(* IEC 61131-3 sources: PortalRobot/Portal_robot/Device/application (part 2) *)

(* ---- PLC_PRG.ReadIoOverrides.st ---- *)
METHOD PRIVATE ReadIoOverrides

// --- BEGIN IMPLEMENTATION ---

udiIoNowMs := TIME_TO_UDINT(TIME());
IF NOT xIoInitialized THEN
    GVL_HMI.udiIoBootCounter := GVL_HMI.udiIoBootCounter + UDINT#1;
    IF GVL_HMI.udiIoBootCounter = UDINT#0 THEN GVL_HMI.udiIoBootCounter := UDINT#1; END_IF;
    udiIoLastTickMs := udiIoNowMs;
    // Старый запрос после перезапуска не должен исполняться сам собой.
    GVL_HMI.udiIoOverrideAckSeq := GVL_HMI.udiIoOverrideCommandSeq;
    GVL_HMI.udiIoEmergencyAckSeq := GVL_HMI.udiIoEmergencyCommandSeq;
END_IF;
IF udiIoNowMs >= udiIoLastTickMs THEN
    uliIoClockMs := uliIoClockMs + UDINT_TO_ULINT(udiIoNowMs - udiIoLastTickMs);
ELSE
    uliIoClockMs := uliIoClockMs + ULINT#4294967296 - UDINT_TO_ULINT(udiIoLastTickMs) + UDINT_TO_ULINT(udiIoNowMs);
END_IF;
udiIoLastTickMs := udiIoNowMs;
GVL_HMI.sIoClockMs := ULINT_TO_STRING(uliIoClockMs);

tonIoOverrideWatchdog(IN := GVL_HMI.udiIoOverrideHeartbeat = udiIoHeartbeatSeen, PT := T#3S);
IF GVL_HMI.udiIoOverrideHeartbeat <> udiIoHeartbeatSeen THEN
    udiIoHeartbeatSeen := GVL_HMI.udiIoOverrideHeartbeat;
END_IF;
IF udiIoNowMs >= GVL_HMI.udiIoOverrideHeartbeatAtMs THEN
    uliIoLeaseAgeMs := UDINT_TO_ULINT(udiIoNowMs) - UDINT_TO_ULINT(GVL_HMI.udiIoOverrideHeartbeatAtMs);
ELSE
    uliIoLeaseAgeMs := ULINT#4294967296 + UDINT_TO_ULINT(udiIoNowMs) - UDINT_TO_ULINT(GVL_HMI.udiIoOverrideHeartbeatAtMs);
END_IF;

xIoBusy := GVL_CELL_MANAGER.Status.xRunning OR GVL_CELL_MANAGER.Status.xBusy
    OR GVL_CELL_MANAGER.Status.xStopPending OR GVL_ROBOT.Status.xBusy
    OR xMotionBusy OR xGroupMotionBusy OR xPointCheckActive OR xPointCheckRequest
    OR xPowerTransitionActive OR SIMULATION_DYNAMICS.xBusy
    OR GVL_HMI.xRobotManualExecute OR GVL_HMI.stRobotCommand.xExecute
    OR GVL_CELL_CONTROL.xStart
    OR (GVL_HMI.udiTwinCommandSeq <> GVL_HMI.udiTwinAckSeq);
// Реальный цикл станка нельзя скрыть подменой его DI.
IF xPhysicalNormal AND GVL_PHYSICAL_IO.xMappingVerified THEN
    xIoBusy := xIoBusy OR GVL_PHYSICAL_IO.xDiMachine1CycleActive
        OR GVL_PHYSICAL_IO.xDiMachine2CycleActive OR GVL_PHYSICAL_IO.xDiMachine3CycleActive;
END_IF;
FOR uiIoIndex := UINT#1 TO UINT#3 DO
    xIoBusy := xIoBusy OR GVL_MACHINE.Status[uiIoIndex].xBusy OR GVL_MACHINE.Status[uiIoIndex].xProcessing
        OR GVL_HMI.axMachineManualHatchOpen[uiIoIndex] OR GVL_HMI.axMachineManualHatchClose[uiIoIndex]
        OR GVL_HMI.axMachineManualHatchUnlock[uiIoIndex] OR GVL_HMI.axMachineManualHatchLock[uiIoIndex]
        OR GVL_HMI.axMachineManualChuckOpen[uiIoIndex] OR GVL_HMI.axMachineManualChuckClose[uiIoIndex]
        OR GVL_HMI.astAxisHmiCommand[uiIoIndex].xJogPositive
        OR GVL_HMI.astAxisHmiCommand[uiIoIndex].xJogNegative
        OR GVL_HMI.astAxisHmiCommand[uiIoIndex].xHome
        OR GVL_HMI.astAxisHmiCommand[uiIoIndex].xMoveAbsolute
        OR GVL_HMI.astAxisHmiCommand[uiIoIndex].xMoveRelative;
END_FOR;
FOR uiIoIndex := UINT#1 TO UINT#2 DO
    xIoBusy := xIoBusy OR GVL_MAGAZINE.astStatus[uiIoIndex].xBusy
        OR GVL_TWO_PALLET.astStatus[uiIoIndex].xBusy;
END_FOR;
// Ручной режим сигналов включается одним запросом. Технологических допусков здесь нет.
xIoManualEndedByOperator := FALSE;
IF xIoManualActive AND (NOT GVL_CELL_CONTROL.xManual OR NOT xHmiConnectionAlive
    OR CONTROLLER_DIAGNOSTICS.Status.xAlarmActive
    OR tonIoOverrideWatchdog.Q OR (uliIoLeaseAgeMs > ULINT#3000)
    OR ((GVL_HMI.udiCellModeCommandSeq <> GVL_HMI.udiCellModeAckSeq) AND NOT GVL_HMI.xCellManualRequest)) THEN
    xIoManualActive := FALSE;
END_IF;
// Прямой ручной слой доступен и при зависших Busy/Processing владельцев.
// Их задания отменяются при передаче управления; xIoBusy остаётся диагностикой
// и условием снятия отдельного программного аварийного останова.
GVL_HMI.xIoManualStartAllowed := GVL_CELL_CONTROL.xManual AND NOT xIoManualActive
    AND NOT CONTROLLER_DIAGNOSTICS.Status.xAlarmActive
    AND NOT ((GVL_HMI.udiCellModeCommandSeq <> GVL_HMI.udiCellModeAckSeq) AND NOT GVL_HMI.xCellManualRequest);
xIoOverrideRejected := FALSE;
udiIoRequestSeq := GVL_HMI.udiIoOverrideCommandSeq;
uiIoRequestAction := GVL_HMI.uiIoOverrideAction;
uiIoRequestIndex := GVL_HMI.uiIoOverrideIndex;
xIoRequestValue := GVL_HMI.xIoOverrideValue;
IF udiIoRequestSeq <> GVL_HMI.udiIoOverrideAckSeq THEN
    IF (uiIoRequestAction = UINT#8) OR (uiIoRequestAction = UINT#9) OR (uiIoRequestAction = UINT#7) THEN
        GVL_HMI.uiIoOverrideResult := UINT#4;
        IF IsHmiCommandFresh(udiIssuedAtMs := GVL_HMI.udiIoOverrideIssuedAtMs) THEN
            GVL_HMI.uiIoOverrideResult := UINT#1;
            IF uiIoRequestAction = UINT#8 THEN
                IF NOT xHmiConnectionAlive OR tonIoOverrideWatchdog.Q OR (uliIoLeaseAgeMs > ULINT#3000) THEN
                    GVL_HMI.uiIoOverrideResult := UINT#4;
                ELSIF xIoManualActive THEN
                    // Повтор входа не перезаписывает уже выбранные ручные уровни.
                    GVL_HMI.uiIoOverrideResult := UINT#1;
                ELSIF GVL_HMI.xIoManualStartAllowed THEN
                    FOR uiIoIndex := UINT#1 TO UINT#50 DO
                        axIoDoForceValue[uiIoIndex] := axIoOutput[uiIoIndex];
                        axIoDoForced[uiIoIndex] := FALSE;
                    END_FOR;
                    xIoManualActive := TRUE;
                ELSE
                    GVL_HMI.uiIoOverrideResult := UINT#2;
                END_IF;
            ELSE
                xIoManualActive := FALSE;
                xIoManualEndedByOperator := TRUE;
            END_IF;
        END_IF;
        // Для входа/выхода из режима Ack выдаёт ApplyIoOutputOverrides после назначения DO.
    END_IF;
END_IF;

GVL_HMI.xIoManualControlActive := xIoManualActive;
GVL_HMI.xIoManualStartAllowed := GVL_HMI.xIoManualStartAllowed AND NOT xIoManualActive;
GVL_HMI.xIoOverrideAllowed := xIoManualActive AND GVL_CELL_CONTROL.xManual;
IF GVL_HMI.xIoOverrideAllowed THEN GVL_HMI.uiIoOverrideBlockReason := UINT#0;
ELSIF NOT GVL_CELL_CONTROL.xManual THEN GVL_HMI.uiIoOverrideBlockReason := UINT#2;
ELSE GVL_HMI.uiIoOverrideBlockReason := UINT#7;
END_IF;

IF NOT GVL_HMI.xIoOverrideAllowed THEN
    FOR uiIoIndex := UINT#1 TO UINT#84 DO
        IF axIoForced[uiIoIndex] THEN
            IF xIoManualEndedByOperator THEN
                AppendIoEvent(usiDirection := USINT#1, uiIndex := uiIoIndex, usiKind := USINT#5,
                    xOld := axIoForceValue[uiIoIndex], xNew := axIoRawDi[uiIoIndex]);
            ELSE
                AppendIoEvent(usiDirection := USINT#1, uiIndex := uiIoIndex, usiKind := USINT#6,
                    xOld := axIoForceValue[uiIoIndex], xNew := axIoRawDi[uiIoIndex]);
            END_IF;
            axIoForced[uiIoIndex] := FALSE;
        END_IF;
    END_FOR;
END_IF;

IF (udiIoRequestSeq <> GVL_HMI.udiIoOverrideAckSeq)
AND NOT ((uiIoRequestAction >= UINT#4) AND (uiIoRequestAction <= UINT#9)) THEN
    GVL_HMI.uiIoOverrideResult := UINT#3;
    IF NOT IsHmiCommandFresh(udiIssuedAtMs := GVL_HMI.udiIoOverrideIssuedAtMs) THEN
        GVL_HMI.uiIoOverrideResult := UINT#4;
    ELSIF uiIoRequestAction = UINT#3 THEN
        FOR uiIoIndex := UINT#1 TO UINT#84 DO
            IF axIoForced[uiIoIndex] THEN
                AppendIoEvent(usiDirection := USINT#1, uiIndex := uiIoIndex, usiKind := USINT#5,
                    xOld := axIoForceValue[uiIoIndex], xNew := axIoRawDi[uiIoIndex]);
                axIoForced[uiIoIndex] := FALSE;
            END_IF;
        END_FOR;
        GVL_HMI.uiIoOverrideResult := UINT#1;
    ELSIF (uiIoRequestIndex >= UINT#1) AND (uiIoRequestIndex <= UINT#84) THEN
        IF uiIoRequestAction = UINT#2 THEN
            IF axIoForced[uiIoRequestIndex] THEN
                AppendIoEvent(usiDirection := USINT#1, uiIndex := uiIoRequestIndex, usiKind := USINT#5,
                    xOld := axIoForceValue[uiIoRequestIndex], xNew := axIoRawDi[uiIoRequestIndex]);
                axIoForced[uiIoRequestIndex] := FALSE;
            END_IF;
            GVL_HMI.uiIoOverrideResult := UINT#1;
        ELSIF uiIoRequestAction = UINT#1 THEN
            IF GVL_HMI.xIoOverrideAllowed THEN
                IF NOT axIoForced[uiIoRequestIndex] OR (axIoForceValue[uiIoRequestIndex] <> xIoRequestValue) THEN
                    AppendIoEvent(usiDirection := USINT#1, uiIndex := uiIoRequestIndex, usiKind := USINT#4,
                        xOld := axPhysicalRaw[uiIoRequestIndex], xNew := xIoRequestValue);
                END_IF;
                axIoForced[uiIoRequestIndex] := TRUE;
                axIoForceValue[uiIoRequestIndex] := xIoRequestValue;
                GVL_HMI.uiIoOverrideResult := UINT#1;
            ELSE
                GVL_HMI.uiIoOverrideResult := UINT#2;
            END_IF;
        END_IF;
    END_IF;
    xIoOverrideRejected := GVL_HMI.uiIoOverrideResult <> UINT#1;
    GVL_HMI.udiIoOverrideAckSeq := udiIoRequestSeq;
END_IF;
FOR uiIoIndex := UINT#1 TO UINT#84 DO
    IF axIoForced[uiIoIndex] THEN axPhysicalRaw[uiIoIndex] := axIoForceValue[uiIoIndex]; END_IF;
END_FOR;

(* ---- PLC_PRG.ReadPhysicalInputs.st ---- *)
METHOD PRIVATE ReadPhysicalInputs

// --- BEGIN IMPLEMENTATION ---

// Единственная страница назначения входов. Сначала фильтры, затем технологические FB.
// Тестовые среды используют модели; сырые входы приводов ГК читает RunGeometryControl.
xPhysicalNormal := GVL_CELL_SETTINGS.eTestEnvironment = E_CELL_TEST_ENVIRONMENT.NORMAL;
GVL_PHYSICAL_IO.xNormalActive := xPhysicalNormal AND GVL_PHYSICAL_IO.xMappingVerified;
xPhysicalInputEnable := GVL_PHYSICAL_IO.xNormalActive;

axPhysicalRaw[1] := GVL_PHYSICAL_IO.xDiMachine1Ready;
axPhysicalRaw[2] := GVL_PHYSICAL_IO.xDiMachine1Alarm;
axPhysicalRaw[3] := GVL_PHYSICAL_IO.xDiMachine1DoorOpen;
axPhysicalRaw[4] := GVL_PHYSICAL_IO.xDiMachine1DoorClosed;
axPhysicalRaw[5] := GVL_PHYSICAL_IO.xDiMachine1HatchLocked;
axPhysicalRaw[6] := GVL_PHYSICAL_IO.xDiMachine1SafetyDoorOpen;
axPhysicalRaw[7] := GVL_PHYSICAL_IO.xDiMachine1SafetyDoorClosed;
axPhysicalRaw[8] := GVL_PHYSICAL_IO.xDiMachine1ChuckClamped;
axPhysicalRaw[9] := GVL_PHYSICAL_IO.xDiMachine1ChuckUnclamped;
axPhysicalRaw[10] := GVL_PHYSICAL_IO.xDiMachine1CycleActive;
axPhysicalRaw[11] := GVL_PHYSICAL_IO.xDiMachine1CycleDone;
axPhysicalRaw[12] := GVL_PHYSICAL_IO.xDiMachine2Ready;
axPhysicalRaw[13] := GVL_PHYSICAL_IO.xDiMachine2Alarm;
axPhysicalRaw[14] := GVL_PHYSICAL_IO.xDiMachine2DoorOpen;
axPhysicalRaw[15] := GVL_PHYSICAL_IO.xDiMachine2DoorClosed;
axPhysicalRaw[16] := GVL_PHYSICAL_IO.xDiMachine2HatchLocked;
axPhysicalRaw[17] := GVL_PHYSICAL_IO.xDiMachine2SafetyDoorOpen;
axPhysicalRaw[18] := GVL_PHYSICAL_IO.xDiMachine2SafetyDoorClosed;
axPhysicalRaw[19] := GVL_PHYSICAL_IO.xDiMachine2ChuckClamped;
axPhysicalRaw[20] := GVL_PHYSICAL_IO.xDiMachine2ChuckUnclamped;
axPhysicalRaw[21] := GVL_PHYSICAL_IO.xDiMachine2CycleActive;
axPhysicalRaw[22] := GVL_PHYSICAL_IO.xDiMachine2CycleDone;
axPhysicalRaw[23] := GVL_PHYSICAL_IO.xDiMachine3Ready;
axPhysicalRaw[24] := GVL_PHYSICAL_IO.xDiMachine3Alarm;
axPhysicalRaw[25] := GVL_PHYSICAL_IO.xDiMachine3DoorOpen;
axPhysicalRaw[26] := GVL_PHYSICAL_IO.xDiMachine3DoorClosed;
axPhysicalRaw[27] := GVL_PHYSICAL_IO.xDiMachine3HatchLocked;
axPhysicalRaw[28] := GVL_PHYSICAL_IO.xDiMachine3SafetyDoorOpen;
axPhysicalRaw[29] := GVL_PHYSICAL_IO.xDiMachine3SafetyDoorClosed;
axPhysicalRaw[30] := GVL_PHYSICAL_IO.xDiMachine3ChuckClamped;
axPhysicalRaw[31] := GVL_PHYSICAL_IO.xDiMachine3ChuckUnclamped;
axPhysicalRaw[32] := GVL_PHYSICAL_IO.xDiMachine3CycleActive;
axPhysicalRaw[33] := GVL_PHYSICAL_IO.xDiMachine3CycleDone;
axPhysicalRaw[34] := GVL_PHYSICAL_IO.xDiGripper1Open;
axPhysicalRaw[35] := GVL_PHYSICAL_IO.xDiGripper1Closed;
axPhysicalRaw[36] := GVL_PHYSICAL_IO.xDiGripper2Open;
axPhysicalRaw[37] := GVL_PHYSICAL_IO.xDiGripper2Closed;
axPhysicalRaw[38] := GVL_PHYSICAL_IO.xDiRotatedToBlank;
axPhysicalRaw[39] := GVL_PHYSICAL_IO.xDiRotatedToDetail;
axPhysicalRaw[40] := GVL_PHYSICAL_IO.xDiCellStartButtonInput;
axPhysicalRaw[41] := GVL_PHYSICAL_IO.xDiCellStopButtonInput;
axPhysicalRaw[42] := GVL_PHYSICAL_IO.xDiCellResetButtonInput;
axPhysicalRaw[43] := GVL_PHYSICAL_IO.xDiEmergencyStopStation1Ok;
axPhysicalRaw[44] := GVL_PHYSICAL_IO.xDiEmergencyStopStation2Ok;
axPhysicalRaw[45] := GVL_PHYSICAL_IO.xDiEmergencyStopStation3Ok;
axPhysicalRaw[46] := GVL_PHYSICAL_IO.xDiEmergencyStopStation4Ok;
axPhysicalRaw[47] := GVL_PHYSICAL_IO.xDiEmergencyStopCabinet1Ok;
axPhysicalRaw[48] := GVL_PHYSICAL_IO.xDiEmergencyStopCabinet2Ok;
axPhysicalRaw[49] := GVL_PHYSICAL_IO.xDiEmergencyStopMpgOk;
axPhysicalRaw[50] := GVL_PHYSICAL_IO.xDiDoor1LockClosed;
axPhysicalRaw[51] := GVL_PHYSICAL_IO.xDiDoor2LockClosed;
axPhysicalRaw[52] := GVL_PHYSICAL_IO.xDiDoor3LockClosed;
axPhysicalRaw[53] := GVL_PHYSICAL_IO.xDiDoor4LockClosed;
axPhysicalRaw[54] := GVL_PHYSICAL_IO.xDiSafetyRelayOkInput;
axPhysicalRaw[55] := GVL_PHYSICAL_IO.xDiPhaseRelayOkInput;
axPhysicalRaw[56] := GVL_PHYSICAL_IO.xDiPressureRelayOkInput;
axPhysicalRaw[57] := GVL_PHYSICAL_IO.xDiMpgAxisXInput;
axPhysicalRaw[58] := GVL_PHYSICAL_IO.xDiMpgAxisYInput;
axPhysicalRaw[59] := GVL_PHYSICAL_IO.xDiMpgAxisZInput;
axPhysicalRaw[60] := GVL_PHYSICAL_IO.xDiMpgMultiplier1Input;
axPhysicalRaw[61] := GVL_PHYSICAL_IO.xDiMpgMultiplier10Input;
axPhysicalRaw[62] := GVL_PHYSICAL_IO.xDiMpgMultiplier100Input;
axPhysicalRaw[63] := GVL_PHYSICAL_IO.xDiMagazine1LockIn;
axPhysicalRaw[64] := GVL_PHYSICAL_IO.xDiMagazine1LockOut;
axPhysicalRaw[65] := GVL_PHYSICAL_IO.xDiMagazine1StopIn;
axPhysicalRaw[66] := GVL_PHYSICAL_IO.xDiMagazine1StopOut;
axPhysicalRaw[67] := GVL_PHYSICAL_IO.xDiMagazine1LiftUp;
axPhysicalRaw[68] := GVL_PHYSICAL_IO.xDiMagazine1LiftDown;
axPhysicalRaw[69] := GVL_PHYSICAL_IO.xDiDoor1UnlockButton;
axPhysicalRaw[70] := GVL_PHYSICAL_IO.xDiDoor2UnlockButton;
axPhysicalRaw[71] := GVL_PHYSICAL_IO.xDiDoor3UnlockButton;
axPhysicalRaw[72] := GVL_PHYSICAL_IO.xDiDoor4UnlockButton;
axPhysicalRaw[73] := GVL_PHYSICAL_IO.xDiMagazine2LockIn;
axPhysicalRaw[74] := GVL_PHYSICAL_IO.xDiMagazine2LockOut;
axPhysicalRaw[75] := GVL_PHYSICAL_IO.xDiMagazine2StopIn;
axPhysicalRaw[76] := GVL_PHYSICAL_IO.xDiMagazine2StopOut;
axPhysicalRaw[77] := GVL_PHYSICAL_IO.xDiMagazine2LiftUp;
axPhysicalRaw[78] := GVL_PHYSICAL_IO.xDiMagazine2LiftDown;

axPhysicalRaw[79] := GVL_PHYSICAL_IO.xDiGk1PartAtEnd;
axPhysicalRaw[80] := GVL_PHYSICAL_IO.xDiGk2PartAtEnd;

axPhysicalRaw[81] := GVL_PHYSICAL_IO.xDiGk1DriveAlarm;
axPhysicalRaw[82] := GVL_PHYSICAL_IO.xDiGk1DriveRunning;
axPhysicalRaw[83] := GVL_PHYSICAL_IO.xDiGk2DriveAlarm;
axPhysicalRaw[84] := GVL_PHYSICAL_IO.xDiGk2DriveRunning;
// Клеммы сохраняются отдельно: ручная подмена не пишет в переменную I/O Mapping.
FOR uiIoIndex := UINT#1 TO UINT#84 DO
    axIoRawDi[uiIoIndex] := axPhysicalRaw[uiIoIndex];
END_FOR;
ReadIoOverrides();
FOR uiIoIndex := UINT#1 TO UINT#84 DO
    IF axIoForced[uiIoIndex] THEN
        axPhysicalRaw[uiIoIndex] := axIoForceValue[uiIoIndex];
    END_IF;
END_FOR;

FOR uiPhysicalInput := 1 TO 80 DO
	tPhysicalRise := GVL_CELL_SETTINGS.tInputFilterRise;
	tPhysicalFall := GVL_CELL_SETTINGS.tInputFilterFall;
	// Срабатывание опасного состояния не задерживается; восстановление фильтруется.
	CASE uiPhysicalInput OF
		2, 13, 24, 41:
			tPhysicalRise := T#0MS;
		1, 3, 4, 5, 6, 7, 8, 9, 12, 14, 15, 16, 17, 18, 19, 20, 23, 25, 26, 27, 28, 29, 30, 31, 34, 35, 36, 37, 38, 39, 43, 44, 45, 46, 47, 48, 49, 50, 51, 52, 53, 54, 55, 56, 63, 64, 65, 66, 67, 68, 73, 74, 75, 76, 77, 78, 79, 80:
			tPhysicalFall := T#0MS;
	END_CASE;
	xPhysicalInputEnable := xPhysicalNormal AND (GVL_PHYSICAL_IO.xMappingVerified OR axIoForced[uiPhysicalInput]);
	afbPhysicalInputFilter[uiPhysicalInput](
		xEnable := xPhysicalInputEnable, xInput := axPhysicalRaw[uiPhysicalInput],
		tRise := tPhysicalRise, tFall := tPhysicalFall);
	axPhysicalFiltered[uiPhysicalInput] := afbPhysicalInputFilter[uiPhysicalInput].xFiltered;
	IF NOT xPhysicalInputEnable THEN
		axPhysicalButtonArmed[uiPhysicalInput] := FALSE;
	ELSIF NOT axPhysicalRaw[uiPhysicalInput] THEN
		axPhysicalButtonArmed[uiPhysicalInput] := TRUE;
	END_IF;
END_FOR;

// Датчики используются FB_GEOMETRY_CONTROL; в NORMAL доступна диагностическая подмена до подтверждения карты.
GVL_PHYSICAL_IO.axGkPartAtEnd[1] := axPhysicalFiltered[79];
GVL_PHYSICAL_IO.axGkPartAtEnd[2] := axPhysicalFiltered[80];

IF xPhysicalNormal THEN
	GVL_MACHINE.astPhysicalInput[1].xReady := axPhysicalFiltered[1];
	GVL_MACHINE.astPhysicalInput[1].xAlarm := axPhysicalFiltered[2];
	GVL_MACHINE.astPhysicalInput[1].xDoorOpen := axPhysicalFiltered[3];
	GVL_MACHINE.astPhysicalInput[1].xDoorClosed := axPhysicalFiltered[4];
	GVL_MACHINE.astPhysicalInput[1].xHatchLocked := axPhysicalFiltered[5];
	GVL_MACHINE.astPhysicalInput[1].xSafetyDoorOpen := axPhysicalFiltered[6];
	GVL_MACHINE.astPhysicalInput[1].xSafetyDoorClosed := axPhysicalFiltered[7];
	GVL_MACHINE.astPhysicalInput[1].xChuckClamped := axPhysicalFiltered[8];
	GVL_MACHINE.astPhysicalInput[1].xChuckUnclamped := axPhysicalFiltered[9];
	GVL_MACHINE.astPhysicalInput[1].xCycleActive := axPhysicalFiltered[10];
	GVL_MACHINE.astPhysicalInput[1].xCycleDone := axPhysicalFiltered[11];
	GVL_MACHINE.astPhysicalInput[2].xReady := axPhysicalFiltered[12];
	GVL_MACHINE.astPhysicalInput[2].xAlarm := axPhysicalFiltered[13];
	GVL_MACHINE.astPhysicalInput[2].xDoorOpen := axPhysicalFiltered[14];
	GVL_MACHINE.astPhysicalInput[2].xDoorClosed := axPhysicalFiltered[15];
	GVL_MACHINE.astPhysicalInput[2].xHatchLocked := axPhysicalFiltered[16];
	GVL_MACHINE.astPhysicalInput[2].xSafetyDoorOpen := axPhysicalFiltered[17];
	GVL_MACHINE.astPhysicalInput[2].xSafetyDoorClosed := axPhysicalFiltered[18];
	GVL_MACHINE.astPhysicalInput[2].xChuckClamped := axPhysicalFiltered[19];
	GVL_MACHINE.astPhysicalInput[2].xChuckUnclamped := axPhysicalFiltered[20];
	GVL_MACHINE.astPhysicalInput[2].xCycleActive := axPhysicalFiltered[21];
	GVL_MACHINE.astPhysicalInput[2].xCycleDone := axPhysicalFiltered[22];
	GVL_MACHINE.astPhysicalInput[3].xReady := axPhysicalFiltered[23];
	GVL_MACHINE.astPhysicalInput[3].xAlarm := axPhysicalFiltered[24];
	GVL_MACHINE.astPhysicalInput[3].xDoorOpen := axPhysicalFiltered[25];
	GVL_MACHINE.astPhysicalInput[3].xDoorClosed := axPhysicalFiltered[26];
	GVL_MACHINE.astPhysicalInput[3].xHatchLocked := axPhysicalFiltered[27];
	GVL_MACHINE.astPhysicalInput[3].xSafetyDoorOpen := axPhysicalFiltered[28];
	GVL_MACHINE.astPhysicalInput[3].xSafetyDoorClosed := axPhysicalFiltered[29];
	GVL_MACHINE.astPhysicalInput[3].xChuckClamped := axPhysicalFiltered[30];
	GVL_MACHINE.astPhysicalInput[3].xChuckUnclamped := axPhysicalFiltered[31];
	GVL_MACHINE.astPhysicalInput[3].xCycleActive := axPhysicalFiltered[32];
	GVL_MACHINE.astPhysicalInput[3].xCycleDone := axPhysicalFiltered[33];
	GVL_PHYSICAL_IO.stGripperFeedback.xGripper1Open := axPhysicalFiltered[34];
	GVL_PHYSICAL_IO.stGripperFeedback.xGripper1Closed := axPhysicalFiltered[35];
	GVL_PHYSICAL_IO.stGripperFeedback.xGripper2Open := axPhysicalFiltered[36];
	GVL_PHYSICAL_IO.stGripperFeedback.xGripper2Closed := axPhysicalFiltered[37];
	GVL_PHYSICAL_IO.stGripperFeedback.xRotatedToBlank := axPhysicalFiltered[38];
	GVL_PHYSICAL_IO.stGripperFeedback.xRotatedToDetail := axPhysicalFiltered[39];
	GVL_CELL_SAFETY_IO.xCellStartButtonInput := axPhysicalFiltered[40] AND axPhysicalButtonArmed[40];
	GVL_CELL_SAFETY_IO.xCellStopButtonInput := axPhysicalFiltered[41];
	GVL_CELL_SAFETY_IO.xCellResetButtonInput := axPhysicalFiltered[42] AND axPhysicalButtonArmed[42];
	GVL_CELL_SAFETY_IO.axEmergencyStopButtonStationInput[1] := NOT axPhysicalFiltered[43];
	GVL_CELL_SAFETY_IO.axEmergencyStopButtonStationInput[2] := NOT axPhysicalFiltered[44];
	GVL_CELL_SAFETY_IO.axEmergencyStopButtonStationInput[3] := NOT axPhysicalFiltered[45];
	GVL_CELL_SAFETY_IO.axEmergencyStopButtonStationInput[4] := NOT axPhysicalFiltered[46];
	GVL_CELL_SAFETY_IO.axEmergencyStopCabinetInput[1] := NOT axPhysicalFiltered[47];
	GVL_CELL_SAFETY_IO.axEmergencyStopCabinetInput[2] := NOT axPhysicalFiltered[48];
	GVL_CELL_SAFETY_IO.xEmergencyStopMpgInput := NOT axPhysicalFiltered[49];
	GVL_CELL_SAFETY_IO.axDoorLockClosedInput[1] := axPhysicalFiltered[50];
	GVL_CELL_SAFETY_IO.axDoorLockClosedInput[2] := axPhysicalFiltered[51];
	GVL_CELL_SAFETY_IO.axDoorLockClosedInput[3] := axPhysicalFiltered[52];
	GVL_CELL_SAFETY_IO.axDoorLockClosedInput[4] := axPhysicalFiltered[53];
	GVL_CELL_SAFETY_IO.xSafetyRelayOkInput := axPhysicalFiltered[54];
	GVL_CELL_SAFETY_IO.xPhaseRelayOkInput := axPhysicalFiltered[55];
	GVL_CELL_SAFETY_IO.xPressureRelayOkInput := axPhysicalFiltered[56];
	GVL_CELL_SAFETY_IO.xMpgAxisXInput := axPhysicalFiltered[57];
	GVL_CELL_SAFETY_IO.xMpgAxisYInput := axPhysicalFiltered[58];
	GVL_CELL_SAFETY_IO.xMpgAxisZInput := axPhysicalFiltered[59];
	GVL_CELL_SAFETY_IO.xMpgMultiplier1Input := axPhysicalFiltered[60];
	GVL_CELL_SAFETY_IO.xMpgMultiplier10Input := axPhysicalFiltered[61];
	GVL_CELL_SAFETY_IO.xMpgMultiplier100Input := axPhysicalFiltered[62];
	GVL_TWO_PALLET.astInput[1].xLockIn := axPhysicalFiltered[63];
	GVL_TWO_PALLET.astInput[1].xLockOut := axPhysicalFiltered[64];
	GVL_TWO_PALLET.astInput[1].xStopIn := axPhysicalFiltered[65];
	GVL_TWO_PALLET.astInput[1].xStopOut := axPhysicalFiltered[66];
	GVL_TWO_PALLET.astInput[1].xLiftUp := axPhysicalFiltered[67];
	GVL_TWO_PALLET.astInput[1].xLiftDown := axPhysicalFiltered[68];
	GVL_CELL_SAFETY_IO.axDoorUnlockButtonInput[1] := axPhysicalFiltered[69] AND axPhysicalButtonArmed[69];
	GVL_CELL_SAFETY_IO.axDoorUnlockButtonInput[2] := axPhysicalFiltered[70] AND axPhysicalButtonArmed[70];
	GVL_CELL_SAFETY_IO.axDoorUnlockButtonInput[3] := axPhysicalFiltered[71] AND axPhysicalButtonArmed[71];
	GVL_CELL_SAFETY_IO.axDoorUnlockButtonInput[4] := axPhysicalFiltered[72] AND axPhysicalButtonArmed[72];
	GVL_TWO_PALLET.astInput[2].xLockIn := axPhysicalFiltered[73];
	GVL_TWO_PALLET.astInput[2].xLockOut := axPhysicalFiltered[74];
	GVL_TWO_PALLET.astInput[2].xStopIn := axPhysicalFiltered[75];
	GVL_TWO_PALLET.astInput[2].xStopOut := axPhysicalFiltered[76];
	GVL_TWO_PALLET.astInput[2].xLiftUp := axPhysicalFiltered[77];
	GVL_TWO_PALLET.astInput[2].xLiftDown := axPhysicalFiltered[78];
	GVL_TWO_PALLET.astInput[1].xIoMapped := GVL_PHYSICAL_IO.xNormalActive;
	GVL_TWO_PALLET.astInput[2].xIoMapped := GVL_PHYSICAL_IO.xNormalActive;
	GVL_MACHINE.astPhysicalInput[1].tRemaining := T#0MS;
	GVL_MACHINE.astPhysicalInput[2].tRemaining := T#0MS;
	GVL_MACHINE.astPhysicalInput[3].tRemaining := T#0MS;
ELSIF xPhysicalWasNormal THEN
	GVL_CELL_SAFETY_IO.xCellStartButtonInput := FALSE;
	GVL_CELL_SAFETY_IO.xCellStopButtonInput := FALSE;
	GVL_CELL_SAFETY_IO.xCellResetButtonInput := FALSE;
	GVL_CELL_SAFETY_IO.axEmergencyStopButtonStationInput[1] := FALSE;
	GVL_CELL_SAFETY_IO.axEmergencyStopButtonStationInput[2] := FALSE;
	GVL_CELL_SAFETY_IO.axEmergencyStopButtonStationInput[3] := FALSE;
	GVL_CELL_SAFETY_IO.axEmergencyStopButtonStationInput[4] := FALSE;
	GVL_CELL_SAFETY_IO.axEmergencyStopCabinetInput[1] := FALSE;
	GVL_CELL_SAFETY_IO.axEmergencyStopCabinetInput[2] := FALSE;
	GVL_CELL_SAFETY_IO.xEmergencyStopMpgInput := FALSE;
	GVL_CELL_SAFETY_IO.axDoorLockClosedInput[1] := TRUE;
	GVL_CELL_SAFETY_IO.axDoorLockClosedInput[2] := TRUE;
	GVL_CELL_SAFETY_IO.axDoorLockClosedInput[3] := TRUE;
	GVL_CELL_SAFETY_IO.axDoorLockClosedInput[4] := TRUE;
	GVL_CELL_SAFETY_IO.xSafetyRelayOkInput := TRUE;
	GVL_CELL_SAFETY_IO.xPhaseRelayOkInput := TRUE;
	GVL_CELL_SAFETY_IO.xPressureRelayOkInput := TRUE;
	GVL_CELL_SAFETY_IO.xMpgAxisXInput := FALSE;
	GVL_CELL_SAFETY_IO.xMpgAxisYInput := FALSE;
	GVL_CELL_SAFETY_IO.xMpgAxisZInput := FALSE;
	GVL_CELL_SAFETY_IO.xMpgMultiplier1Input := FALSE;
	GVL_CELL_SAFETY_IO.xMpgMultiplier10Input := FALSE;
	GVL_CELL_SAFETY_IO.xMpgMultiplier100Input := FALSE;
	GVL_CELL_SAFETY_IO.axDoorUnlockButtonInput[1] := FALSE;
	GVL_CELL_SAFETY_IO.axDoorUnlockButtonInput[2] := FALSE;
	GVL_CELL_SAFETY_IO.axDoorUnlockButtonInput[3] := FALSE;
	GVL_CELL_SAFETY_IO.axDoorUnlockButtonInput[4] := FALSE;
END_IF;
xPhysicalWasNormal := xPhysicalNormal;

(* ---- PLC_PRG.RecordIoDiagnostics.st ---- *)
METHOD PRIVATE RecordIoDiagnostics

// --- BEGIN IMPLEMENTATION ---

// Seqlock закрывает весь снимок, включая упаковку масок после добавления событий.
GVL_HMI.udiIoJournalRevision := GVL_HMI.udiIoJournalRevision + UDINT#1;
xIoSnapshotPublishing := TRUE;

axIoOutput[1] := GVL_PHYSICAL_IO.xDoMachine1HatchClosed;
axIoOutput[2] := GVL_PHYSICAL_IO.xDoMachine1HatchUnLock;
axIoOutput[3] := GVL_PHYSICAL_IO.xDoMachine1ClampChuck;
axIoOutput[4] := GVL_PHYSICAL_IO.xDoMachine1UnclampChuck;
axIoOutput[5] := GVL_PHYSICAL_IO.xDoMachine1StartCycle;
axIoOutput[6] := GVL_PHYSICAL_IO.xDoMachine2HatchClosed;
axIoOutput[7] := GVL_PHYSICAL_IO.xDoMachine2HatchUnLock;
axIoOutput[8] := GVL_PHYSICAL_IO.xDoMachine2ClampChuck;
axIoOutput[9] := GVL_PHYSICAL_IO.xDoMachine2UnclampChuck;
axIoOutput[10] := GVL_PHYSICAL_IO.xDoMachine2StartCycle;
axIoOutput[11] := GVL_PHYSICAL_IO.xDoMachine3HatchClosed;
axIoOutput[12] := GVL_PHYSICAL_IO.xDoMachine3HatchUnLock;
axIoOutput[13] := GVL_PHYSICAL_IO.xDoMachine3ClampChuck;
axIoOutput[14] := GVL_PHYSICAL_IO.xDoMachine3UnclampChuck;
axIoOutput[15] := GVL_PHYSICAL_IO.xDoMachine3StartCycle;
axIoOutput[16] := GVL_PHYSICAL_IO.xDoGripper1Open;
axIoOutput[17] := GVL_PHYSICAL_IO.xDoGripper2Open;
axIoOutput[18] := GVL_PHYSICAL_IO.xDoRotateToDetail;
axIoOutput[19] := GVL_PHYSICAL_IO.xDoDoor1Unlock;
axIoOutput[27] := GVL_PHYSICAL_IO.xDoDoor1ButtonLamp;
axIoOutput[20] := GVL_PHYSICAL_IO.xDoDoor2Unlock;
axIoOutput[28] := GVL_PHYSICAL_IO.xDoDoor2ButtonLamp;
axIoOutput[21] := GVL_PHYSICAL_IO.xDoDoor3Unlock;
axIoOutput[29] := GVL_PHYSICAL_IO.xDoDoor3ButtonLamp;
axIoOutput[22] := GVL_PHYSICAL_IO.xDoDoor4Unlock;
axIoOutput[30] := GVL_PHYSICAL_IO.xDoDoor4ButtonLamp;
axIoOutput[23] := GVL_PHYSICAL_IO.xDoSafetyRelayReset;
axIoOutput[24] := GVL_PHYSICAL_IO.xDoSignalTowerGreenOutput;
axIoOutput[25] := GVL_PHYSICAL_IO.xDoSignalTowerAmberOutput;
axIoOutput[26] := GVL_PHYSICAL_IO.xDoSignalTowerRedOutput;
axIoOutput[31] := GVL_PHYSICAL_IO.xDoMagazine1LockIn;
axIoOutput[32] := GVL_PHYSICAL_IO.xDoMagazine1LockOut;
axIoOutput[33] := GVL_PHYSICAL_IO.xDoMagazine1StopIn;
axIoOutput[34] := GVL_PHYSICAL_IO.xDoMagazine1StopOut;
axIoOutput[35] := GVL_PHYSICAL_IO.xDoMagazine1LiftUp;
axIoOutput[36] := GVL_PHYSICAL_IO.xDoMagazine1LiftDown;
axIoOutput[43] := GVL_PHYSICAL_IO.xDoMagazine2LockIn;
axIoOutput[44] := GVL_PHYSICAL_IO.xDoMagazine2LockOut;
axIoOutput[45] := GVL_PHYSICAL_IO.xDoMagazine2StopIn;
axIoOutput[46] := GVL_PHYSICAL_IO.xDoMagazine2StopOut;
axIoOutput[47] := GVL_PHYSICAL_IO.xDoMagazine2LiftUp;
axIoOutput[48] := GVL_PHYSICAL_IO.xDoMagazine2LiftDown;
axIoOutput[37] := FALSE; // Удалённый сигнал; индекс журнала не переиспользовать.
axIoOutput[38] := FALSE; // Удалённый сигнал; индекс журнала не переиспользовать.
axIoOutput[39] := FALSE; // Удалённый сигнал; индекс журнала не переиспользовать.
axIoOutput[40] := GVL_PHYSICAL_IO.xDoCellAlarmHorn;
axIoOutput[41] := GVL_PHYSICAL_IO.xDoGk1DriveRun;
axIoOutput[42] := GVL_PHYSICAL_IO.xDoGk1DriveReset;
axIoOutput[49] := GVL_PHYSICAL_IO.xDoGk2DriveRun;
axIoOutput[50] := GVL_PHYSICAL_IO.xDoGk2DriveReset;
FOR uiIoIndex := UINT#1 TO UINT#80 DO
    axIoUsedDi[uiIoIndex] := axPhysicalFiltered[uiIoIndex];
END_FOR;
FOR uiIoIndex := UINT#81 TO UINT#84 DO
    axIoUsedDi[uiIoIndex] := xPhysicalNormal AND (GVL_PHYSICAL_IO.xMappingVerified OR axIoForced[uiIoIndex]) AND axPhysicalRaw[uiIoIndex];
END_FOR;
FOR uiIoIndex := UINT#1 TO UINT#84 DO
    IF xIoInitialized AND (axIoRawDi[uiIoIndex] <> axIoPreviousRaw[uiIoIndex]) THEN
        AppendIoEvent(usiDirection := USINT#1, uiIndex := uiIoIndex, usiKind := USINT#1,
            xOld := axIoPreviousRaw[uiIoIndex], xNew := axIoRawDi[uiIoIndex]);
    END_IF;
    IF xIoInitialized AND (axIoUsedDi[uiIoIndex] <> axIoPreviousUsed[uiIoIndex]) THEN
        AppendIoEvent(usiDirection := USINT#1, uiIndex := uiIoIndex, usiKind := USINT#2,
            xOld := axIoPreviousUsed[uiIoIndex], xNew := axIoUsedDi[uiIoIndex]);
    END_IF;
    axIoPreviousRaw[uiIoIndex] := axIoRawDi[uiIoIndex];
    axIoPreviousUsed[uiIoIndex] := axIoUsedDi[uiIoIndex];
END_FOR;
FOR uiIoIndex := UINT#1 TO UINT#50 DO
    IF xIoInitialized AND ((uiIoIndex < UINT#37) OR (uiIoIndex > UINT#39)) AND (axIoOutput[uiIoIndex] <> axIoPreviousOutput[uiIoIndex]) THEN
        AppendIoEvent(usiDirection := USINT#2, uiIndex := uiIoIndex, usiKind := USINT#3,
            xOld := axIoPreviousOutput[uiIoIndex], xNew := axIoOutput[uiIoIndex]);
    END_IF;
    axIoPreviousOutput[uiIoIndex] := axIoOutput[uiIoIndex];
END_FOR;
xIoInitialized := TRUE; // Первый снимок — начальный уровень, а не 131 выдуманное переключение.

FOR uiIoWord := UINT#1 TO UINT#3 DO
    GVL_HMI.adwIoRawDi[uiIoWord] := DWORD#0;
    GVL_HMI.adwIoUsedDi[uiIoWord] := DWORD#0;
    GVL_HMI.adwIoForcedDi[uiIoWord] := DWORD#0;
END_FOR;
FOR uiIoWord := UINT#1 TO UINT#2 DO
    GVL_HMI.adwIoDo[uiIoWord] := DWORD#0;
    GVL_HMI.adwIoDoAllowed[uiIoWord] := DWORD#0;
    GVL_HMI.adwIoDoOnAllowed[uiIoWord] := DWORD#0;
    GVL_HMI.adwIoForcedDo[uiIoWord] := DWORD#0;
    GVL_HMI.adwIoInhibitedDo[uiIoWord] := DWORD#0;
END_FOR;
GVL_HMI.uiIoForcedCount := UINT#0;
FOR uiIoIndex := UINT#1 TO UINT#84 DO
    uiIoWord := ((uiIoIndex - UINT#1) / UINT#32) + UINT#1;
    uiIoBit := (uiIoIndex - UINT#1) MOD UINT#32;
    dwIoBit := SHL(DWORD#1, uiIoBit);
    IF axIoRawDi[uiIoIndex] THEN GVL_HMI.adwIoRawDi[uiIoWord] := GVL_HMI.adwIoRawDi[uiIoWord] OR dwIoBit; END_IF;
    IF axIoUsedDi[uiIoIndex] THEN GVL_HMI.adwIoUsedDi[uiIoWord] := GVL_HMI.adwIoUsedDi[uiIoWord] OR dwIoBit; END_IF;
    IF axIoForced[uiIoIndex] THEN
        GVL_HMI.adwIoForcedDi[uiIoWord] := GVL_HMI.adwIoForcedDi[uiIoWord] OR dwIoBit;
        GVL_HMI.uiIoForcedCount := GVL_HMI.uiIoForcedCount + UINT#1;
    END_IF;
END_FOR;
FOR uiIoIndex := UINT#1 TO UINT#50 DO
    uiIoWord := ((uiIoIndex - UINT#1) / UINT#32) + UINT#1;
    uiIoBit := (uiIoIndex - UINT#1) MOD UINT#32;
    dwIoBit := SHL(DWORD#1, uiIoBit);
    IF axIoDoAllowed[uiIoIndex] THEN GVL_HMI.adwIoDoAllowed[uiIoWord] := GVL_HMI.adwIoDoAllowed[uiIoWord] OR dwIoBit; END_IF;
    IF axIoDoOnAllowed[uiIoIndex] THEN GVL_HMI.adwIoDoOnAllowed[uiIoWord] := GVL_HMI.adwIoDoOnAllowed[uiIoWord] OR dwIoBit; END_IF;
    IF axIoDoForced[uiIoIndex] THEN GVL_HMI.adwIoForcedDo[uiIoWord] := GVL_HMI.adwIoForcedDo[uiIoWord] OR dwIoBit; END_IF;
    IF axIoDoInhibited[uiIoIndex] THEN GVL_HMI.adwIoInhibitedDo[uiIoWord] := GVL_HMI.adwIoInhibitedDo[uiIoWord] OR dwIoBit; END_IF;
    IF axIoOutput[uiIoIndex] THEN GVL_HMI.adwIoDo[uiIoWord] := GVL_HMI.adwIoDo[uiIoWord] OR SHL(DWORD#1, uiIoBit); END_IF;
END_FOR;
xIoSnapshotPublishing := FALSE;
GVL_HMI.udiIoJournalRevision := GVL_HMI.udiIoJournalRevision + UDINT#1;

(* ---- PLC_PRG.ResetIoEmergencyStop.st ---- *)
METHOD PRIVATE ResetIoEmergencyStop

// --- BEGIN IMPLEMENTATION ---

// Сырые аппаратные сигналы используются для снятия программного останова.
// Прямое ручное I/O этим условием не блокируется.
xIoRawSafetyOk := GVL_PHYSICAL_IO.xMappingVerified
    AND GVL_PHYSICAL_IO.xDiEmergencyStopStation1Ok
    AND GVL_PHYSICAL_IO.xDiEmergencyStopStation2Ok
    AND GVL_PHYSICAL_IO.xDiEmergencyStopStation3Ok
    AND GVL_PHYSICAL_IO.xDiEmergencyStopStation4Ok
    AND GVL_PHYSICAL_IO.xDiEmergencyStopCabinet1Ok
    AND GVL_PHYSICAL_IO.xDiEmergencyStopCabinet2Ok
    AND GVL_PHYSICAL_IO.xDiEmergencyStopMpgOk
    AND GVL_PHYSICAL_IO.xDiSafetyRelayOkInput
    AND GVL_PHYSICAL_IO.xDiPhaseRelayOkInput
    AND GVL_PHYSICAL_IO.xDiPressureRelayOkInput;
// Снять программный останов можно только после останова. Снятие не запускает механизм.
GVL_HMI.xIoEmergencyResetAllowed := GVL_HMI.xIoEmergencyStopActive
    AND GVL_CELL_CONTROL.xManual AND NOT xIoBusy AND xHmiConnectionAlive
    AND CELL_SAFETY.Status.xReady
    AND ((GVL_CELL_SETTINGS.eTestEnvironment <> E_CELL_TEST_ENVIRONMENT.NORMAL) OR xIoRawSafetyOk);
IF GVL_HMI.xIoEmergencyStopActive THEN
    GVL_CELL_CONTROL.xStart := FALSE;
    GVL_CELL_CONTROL.xEnable := FALSE;
    GVL_CELL_CONTROL.xManual := TRUE;
    xRobotHmiPermit := FALSE;
END_IF;
IF xIoEmergencyResetRequested THEN
    GVL_HMI.uiIoEmergencyResult := UINT#3;
    IF NOT IsHmiCommandFresh(udiIssuedAtMs := GVL_HMI.udiIoEmergencyIssuedAtMs) THEN
        GVL_HMI.uiIoEmergencyResult := UINT#4;
    ELSIF GVL_HMI.uiIoEmergencyAction = UINT#2 THEN
        IF GVL_HMI.xIoEmergencyResetAllowed THEN
            GVL_HMI.xIoEmergencyStopActive := FALSE;
            GVL_HMI.uiIoEmergencyResult := UINT#1;
        ELSE GVL_HMI.uiIoEmergencyResult := UINT#2;
        END_IF;
    END_IF;
    xIoEmergencyResetRejected := GVL_HMI.uiIoEmergencyResult <> UINT#1;
    GVL_HMI.udiIoEmergencyAckSeq := udiIoEmergencyRequestSeq;
END_IF;

(* ---- PLC_PRG.RunAlarms.st ---- *)
METHOD PRIVATE RunAlarms

// --- BEGIN IMPLEMENTATION ---

// Единая кнопка подсвечивается только тогда, когда существует хотя бы одна авария
// и каждый активный владелец общей команды готов принять тот же импульс сброса.
// Диагностические защёлки симуляторов станков сюда не входят: они обслуживаются
// отдельной командой «Сброс симулятора» на экране инъекций.
xAlarmResetRequired := CONTROLLER_DIAGNOSTICS.Status.xAlarmActive
    OR (GVL_GEOMETRY_CONTROL.xSupported AND (GVL_GEOMETRY_CONTROL.astStatus[1].xError
	OR GVL_GEOMETRY_CONTROL.astStatus[2].xError))
	OR GVL_CELL_MANAGER.Status.xError
	OR (CELL_SAFETY.Error.dwAlarmActive <> DWORD#0)
	OR GVL_ROBOT.Status.xError
	OR GVL_MACHINE.Status[1].xError
	OR GVL_MACHINE.Status[2].xError
	OR GVL_MACHINE.Status[3].xError
	OR GVL_MAGAZINE.astStatus[1].xError
	OR GVL_MAGAZINE.astStatus[2].xError
	OR (NOT GVL_HMI.xModbusMode AND GVL_AXIS.arrAxis[1].Status.xError)
	OR (NOT GVL_HMI.xModbusMode AND GVL_AXIS.arrAxis[2].Status.xError)
	OR (NOT GVL_HMI.xModbusMode AND GVL_AXIS.arrAxis[3].Status.xError)
	OR (NOT GVL_HMI.xModbusMode AND GVL_AXIS_GROUP.AxisGroup.Status.xLocalError)
	OR (NOT GVL_HMI.xModbusMode AND GVL_AXIS_GROUP.AxisGroup.Status.xLogicalError)
	OR (NOT GVL_HMI.xModbusMode AND GVL_AXIS_GROUP.AxisGroup.Status.xGroupError)
	OR (NOT GVL_HMI.xModbusMode AND (GVL_MOTION_MANAGER.stMotionManager.Error.dwAlarmActive <> DWORD#0))
	OR (NOT GVL_HMI.xModbusMode AND (GVL_POINT_MANAGER.PointManager.Error.dwAlarmActive <> DWORD#0))
	OR (NOT GVL_HMI.xModbusMode AND (GVL_ROBOT.GripperError.dwAlarmActive <> DWORD#0));

xAlarmResetAllowed := ((GVL_TWO_PALLET.uiMode = 0) OR ((NOT GVL_TWO_PALLET.astStatus[1].xError OR GVL_TWO_PALLET.astStatus[1].xResetAllowed) AND (NOT GVL_TWO_PALLET.astStatus[2].xError OR GVL_TWO_PALLET.astStatus[2].xResetAllowed))) AND xAlarmResetRequired
	AND (CELL_SAFETY.Error.dwAlarmActive = DWORD#0)
    AND (NOT CONTROLLER_DIAGNOSTICS.Status.xAlarmActive OR CONTROLLER_DIAGNOSTICS.Status.xResetAllowed)
	AND (NOT GVL_GEOMETRY_CONTROL.xSupported OR NOT GVL_GEOMETRY_CONTROL.astStatus[1].xError OR GVL_GEOMETRY_CONTROL.astStatus[1].xResetAllowed)
	AND (NOT GVL_GEOMETRY_CONTROL.xSupported OR NOT GVL_GEOMETRY_CONTROL.astStatus[2].xError OR GVL_GEOMETRY_CONTROL.astStatus[2].xResetAllowed)
	AND (NOT GVL_CELL_MANAGER.Status.xError OR GVL_CELL_MANAGER.Status.xResetAllowed)
	AND (NOT GVL_ROBOT.Status.xError OR GVL_ROBOT.Status.xResetAllowed)
	AND (NOT GVL_MACHINE.Status[1].xError OR GVL_MACHINE.Status[1].xResetAllowed)
	AND (NOT GVL_MACHINE.Status[2].xError OR GVL_MACHINE.Status[2].xResetAllowed)
	AND (NOT GVL_MACHINE.Status[3].xError OR GVL_MACHINE.Status[3].xResetAllowed)
	AND (NOT GVL_MAGAZINE.astPartStatus[1].xError
		OR (GVL_MAGAZINE.astError[1].dwAlarmActive = DWORD#0)
		OR fbMagazine1.FaultStatus.xResetAllowed)
	AND (NOT GVL_MAGAZINE.astPartStatus[2].xError
		OR (GVL_MAGAZINE.astError[2].dwAlarmActive = DWORD#0)
		OR fbMagazine2.FaultStatus.xResetAllowed)
	AND (GVL_HMI.xModbusMode OR NOT GVL_AXIS.arrAxis[1].Status.xError OR AXIS_X.FaultStatus.xResetAllowed)
	AND (GVL_HMI.xModbusMode OR NOT GVL_AXIS.arrAxis[2].Status.xError OR AXIS_Y.FaultStatus.xResetAllowed)
	AND (GVL_HMI.xModbusMode OR NOT GVL_AXIS.arrAxis[3].Status.xError OR AXIS_Z.FaultStatus.xResetAllowed)
	AND (GVL_HMI.xModbusMode OR NOT (GVL_AXIS_GROUP.AxisGroup.Status.xLocalError
		OR GVL_AXIS_GROUP.AxisGroup.Status.xLogicalError
		OR GVL_AXIS_GROUP.AxisGroup.Status.xGroupError)
		OR GROUP_XYZ.FaultStatus.xResetAllowed)
	AND (GVL_HMI.xModbusMode OR (GVL_MOTION_MANAGER.stMotionManager.Error.dwAlarmActive = DWORD#0)
		OR GVL_ROBOT.Status.xResetAllowed)
	AND (GVL_HMI.xModbusMode OR (GVL_POINT_MANAGER.PointManager.Error.dwAlarmActive = DWORD#0)
		OR (GVL_ROBOT.Status.xResetAllowed AND ROBOT.FaultStatus.stPoint.xResetAllowed))
	AND (GVL_HMI.xModbusMode OR (GVL_ROBOT.GripperError.dwAlarmActive = DWORD#0)
		OR (GVL_ROBOT.Status.xResetAllowed AND ROBOT.FaultStatus.stGripper.xResetAllowed));

// Два владельца предупреждений используют один источник журнала и общий счётчик.
FOR uiTwin := 1 TO 2 DO
	IF GVL_MAGAZINE.astDiag[uiTwin].stWarning.udiSequence <> audiPartWarningSeen[uiTwin] THEN
		audiPartWarningSeen[uiTwin] := GVL_MAGAZINE.astDiag[uiTwin].stWarning.udiSequence;
		astMagazineWarningMerged[uiTwin].uiCode := GVL_MAGAZINE.astDiag[uiTwin].stWarning.uiCode;
		astMagazineWarningMerged[uiTwin].udiSequence := astMagazineWarningMerged[uiTwin].udiSequence + 1;
	END_IF;
	IF GVL_TWO_PALLET.astDiag[uiTwin].stWarning.udiSequence <> audiTwinWarningSeen[uiTwin] THEN
		audiTwinWarningSeen[uiTwin] := GVL_TWO_PALLET.astDiag[uiTwin].stWarning.udiSequence;
		astMagazineWarningMerged[uiTwin].uiCode := GVL_TWO_PALLET.astDiag[uiTwin].stWarning.uiCode;
		astMagazineWarningMerged[uiTwin].udiSequence := astMagazineWarningMerged[uiTwin].udiSequence + 1;
	END_IF;
END_FOR;

// В журнал передаются все активные ошибки и предупреждения каждого функционального блока.
astAlarmSource[18].eSource := E_ALARM_SOURCE.GEOMETRY_1;
astAlarmSource[19].eSource := E_ALARM_SOURCE.GEOMETRY_2;
FOR uiGeometry := UINT#1 TO UINT#2 DO
	IF GVL_GEOMETRY_CONTROL.xSupported THEN
		astAlarmSource[17 + uiGeometry].dwAlarmActive := GVL_GEOMETRY_CONTROL.astActiveMemory[uiGeometry].dwAlarm;
	ELSE astAlarmSource[17 + uiGeometry].dwAlarmActive := DWORD#0; END_IF;
	astAlarmSource[17 + uiGeometry].xRobotStopRequired := GVL_GEOMETRY_CONTROL.astStatus[uiGeometry].xRobotStopRequired;
	astAlarmSource[17 + uiGeometry].xGlobalError := GVL_CELL_CONTROL.xGlobalError;
	astAlarmSource[17 + uiGeometry].stWarning := GVL_GEOMETRY_CONTROL.astWarning[uiGeometry];
END_FOR;
astAlarmSource[1].eSource := E_ALARM_SOURCE.CELL;
astAlarmSource[1].dwAlarmActive := GVL_CELL_MANAGER.Error.dwAlarmActive;
astAlarmSource[1].xRobotStopRequired := FALSE;
astAlarmSource[1].xGlobalError := GVL_CELL_CONTROL.xGlobalError;
astAlarmSource[1].stWarning := GVL_CELL_MANAGER.Diag.stWarning;

// Каждый владелец сохраняет собственные код и счётчик. Подмена Diag ячейки
// чужим событием приводила к откату на старое предупреждение в следующем скане.
// ALARM_MANAGER регистрирует все три канала независимо под источником CELL.
astAdditionalCellWarning[1] := GVL_MULTI_TYPE.ConfigStatus.stWarning;
astAdditionalCellWarning[2] := GVL_GEOMETRY_CONTROL.stCellWarning;

astAlarmSource[2].eSource := E_ALARM_SOURCE.ROBOT;
astAlarmSource[2].dwAlarmActive := GVL_ROBOT.Error.dwAlarmActive;
astAlarmSource[2].xRobotStopRequired := FALSE;
astAlarmSource[2].xGlobalError := GVL_CELL_CONTROL.xGlobalError;
astAlarmSource[2].stWarning := GVL_ROBOT.Diag.stWarning;

astAlarmSource[3].eSource := E_ALARM_SOURCE.MACHINE_1;
astAlarmSource[3].dwAlarmActive := GVL_MACHINE.Error[1].dwAlarmActive;
astAlarmSource[3].xRobotStopRequired := GVL_MACHINE.Status[1].xCriticalError;
astAlarmSource[3].xGlobalError := GVL_CELL_CONTROL.xGlobalError;
astAlarmSource[3].stWarning := GVL_MACHINE.Diag[1].stWarning;

astAlarmSource[4].eSource := E_ALARM_SOURCE.MACHINE_2;
astAlarmSource[4].dwAlarmActive := GVL_MACHINE.Error[2].dwAlarmActive;
astAlarmSource[4].xRobotStopRequired := GVL_MACHINE.Status[2].xCriticalError;
astAlarmSource[4].xGlobalError := GVL_CELL_CONTROL.xGlobalError;
astAlarmSource[4].stWarning := GVL_MACHINE.Diag[2].stWarning;

astAlarmSource[5].eSource := E_ALARM_SOURCE.MACHINE_3;
astAlarmSource[5].dwAlarmActive := GVL_MACHINE.Error[3].dwAlarmActive;
astAlarmSource[5].xRobotStopRequired := GVL_MACHINE.Status[3].xCriticalError;
astAlarmSource[5].xGlobalError := GVL_CELL_CONTROL.xGlobalError;
astAlarmSource[5].stWarning := GVL_MACHINE.Diag[3].stWarning;

astAlarmSource[6].eSource := E_ALARM_SOURCE.MAGAZINE_LOGIC_1;
astAlarmSource[6].dwAlarmActive := GVL_MAGAZINE.astError[1].dwAlarmActive;
astAlarmSource[6].xRobotStopRequired := GVL_MAGAZINE.astStatus[1].xRobotStopRequired;
astAlarmSource[6].xGlobalError := GVL_CELL_CONTROL.xGlobalError;
astAlarmSource[6].stWarning := astMagazineWarningMerged[1];

astAlarmSource[7].eSource := E_ALARM_SOURCE.MAGAZINE_LOGIC_2;
astAlarmSource[7].dwAlarmActive := GVL_MAGAZINE.astError[2].dwAlarmActive;
astAlarmSource[7].xRobotStopRequired := GVL_MAGAZINE.astStatus[2].xRobotStopRequired;
astAlarmSource[7].xGlobalError := GVL_CELL_CONTROL.xGlobalError;
astAlarmSource[7].stWarning := astMagazineWarningMerged[2];

// Числовые коды 7 и 8 зарезервированы, чтобы старые записи SQLite не начали
// отображаться как аварии осей X/Y после удаления приводов магазинов.
astAlarmSource[8].eSource := E_ALARM_SOURCE.RESERVED_LEGACY_MAGAZINE_AXIS_1;
astAlarmSource[8].dwAlarmActive := DWORD#0;
astAlarmSource[8].xRobotStopRequired := FALSE;
astAlarmSource[8].xGlobalError := GVL_CELL_CONTROL.xGlobalError;
astAlarmSource[8].stWarning.uiCode := UINT#0;
astAlarmSource[8].stWarning.udiSequence := UDINT#0;

astAlarmSource[9].eSource := E_ALARM_SOURCE.RESERVED_LEGACY_MAGAZINE_AXIS_2;
astAlarmSource[9].dwAlarmActive := DWORD#0;
astAlarmSource[9].xRobotStopRequired := FALSE;
astAlarmSource[9].xGlobalError := GVL_CELL_CONTROL.xGlobalError;
astAlarmSource[9].stWarning.uiCode := UINT#0;
astAlarmSource[9].stWarning.udiSequence := UDINT#0;

astAlarmSource[10].eSource := E_ALARM_SOURCE.AXIS_X;
IF GVL_HMI.xModbusMode THEN astAlarmSource[10].dwAlarmActive := DWORD#0;
ELSE astAlarmSource[10].dwAlarmActive := GVL_AXIS.arrAxis[1].Error.dwAlarmActive; END_IF;
astAlarmSource[10].xRobotStopRequired := FALSE;
astAlarmSource[10].xGlobalError := GVL_CELL_CONTROL.xGlobalError;
astAlarmSource[10].stWarning := GVL_AXIS.arrAxis[1].Diag.stWarning;

astAlarmSource[11].eSource := E_ALARM_SOURCE.AXIS_Y;
IF GVL_HMI.xModbusMode THEN astAlarmSource[11].dwAlarmActive := DWORD#0;
ELSE astAlarmSource[11].dwAlarmActive := GVL_AXIS.arrAxis[2].Error.dwAlarmActive; END_IF;
astAlarmSource[11].xRobotStopRequired := FALSE;
astAlarmSource[11].xGlobalError := GVL_CELL_CONTROL.xGlobalError;
astAlarmSource[11].stWarning := GVL_AXIS.arrAxis[2].Diag.stWarning;

astAlarmSource[12].eSource := E_ALARM_SOURCE.AXIS_Z;
IF GVL_HMI.xModbusMode THEN astAlarmSource[12].dwAlarmActive := DWORD#0;
ELSE astAlarmSource[12].dwAlarmActive := GVL_AXIS.arrAxis[3].Error.dwAlarmActive; END_IF;
astAlarmSource[12].xRobotStopRequired := FALSE;
astAlarmSource[12].xGlobalError := GVL_CELL_CONTROL.xGlobalError;
astAlarmSource[12].stWarning := GVL_AXIS.arrAxis[3].Diag.stWarning;

astAlarmSource[13].eSource := E_ALARM_SOURCE.AXIS_GROUP;
IF GVL_HMI.xModbusMode THEN astAlarmSource[13].dwAlarmActive := DWORD#0;
ELSE astAlarmSource[13].dwAlarmActive := GVL_AXIS_GROUP.AxisGroup.Error.dwAlarmActive; END_IF;
astAlarmSource[13].xRobotStopRequired := FALSE;
astAlarmSource[13].xGlobalError := GVL_CELL_CONTROL.xGlobalError;
astAlarmSource[13].stWarning := GVL_AXIS_GROUP.AxisGroup.Diag.stWarning;

astAlarmSource[14].eSource := E_ALARM_SOURCE.MOTION_MANAGER;
IF GVL_HMI.xModbusMode THEN astAlarmSource[14].dwAlarmActive := DWORD#0;
ELSE astAlarmSource[14].dwAlarmActive := GVL_MOTION_MANAGER.stMotionManager.Error.dwAlarmActive; END_IF;
astAlarmSource[14].xRobotStopRequired := FALSE;
astAlarmSource[14].xGlobalError := GVL_CELL_CONTROL.xGlobalError;
astAlarmSource[14].stWarning := GVL_MOTION_MANAGER.stMotionManager.Diag.stWarning;

astAlarmSource[15].eSource := E_ALARM_SOURCE.POINT_MANAGER;
IF GVL_HMI.xModbusMode THEN astAlarmSource[15].dwAlarmActive := DWORD#0;
ELSE astAlarmSource[15].dwAlarmActive := GVL_POINT_MANAGER.PointManager.Error.dwAlarmActive; END_IF;
astAlarmSource[15].xRobotStopRequired := FALSE;
astAlarmSource[15].xGlobalError := GVL_CELL_CONTROL.xGlobalError;
astAlarmSource[15].stWarning := GVL_POINT_MANAGER.PointManager.Diag.stWarning;

astAlarmSource[16].eSource := E_ALARM_SOURCE.GRIPPER;
IF GVL_HMI.xModbusMode THEN astAlarmSource[16].dwAlarmActive := DWORD#0;
ELSE astAlarmSource[16].dwAlarmActive := GVL_ROBOT.GripperError.dwAlarmActive; END_IF;
astAlarmSource[16].xRobotStopRequired := FALSE;
astAlarmSource[16].xGlobalError := GVL_CELL_CONTROL.xGlobalError;
astAlarmSource[16].stWarning := GVL_ROBOT.GripperDiag.stWarning;

astAlarmSource[17].eSource := E_ALARM_SOURCE.CELL_SAFETY;
astAlarmSource[17].dwAlarmActive := CELL_SAFETY.Error.dwAlarmActive;
astAlarmSource[17].xRobotStopRequired := TRUE;
astAlarmSource[17].xGlobalError := CELL_SAFETY.Status.xGlobalError;
astAlarmSource[17].stWarning := CELL_SAFETY.Diag.stWarning;

astAlarmSource[20].eSource := E_ALARM_SOURCE.CONTROLLER_CPU_1;
astAlarmSource[20].dwAlarmActive := CONTROLLER_DIAGNOSTICS.Status.dwCpuAlarm1;
astAlarmSource[20].xGlobalError := TRUE;
astAlarmSource[20].stWarning := CONTROLLER_DIAGNOSTICS.stWarning;
astAlarmSource[21].eSource := E_ALARM_SOURCE.CONTROLLER_CPU_2;
astAlarmSource[21].dwAlarmActive := CONTROLLER_DIAGNOSTICS.Status.dwCpuAlarm2;
astAlarmSource[21].xGlobalError := TRUE;
astAlarmSource[22].eSource := E_ALARM_SOURCE.CONTROLLER_MODULES;
astAlarmSource[22].dwAlarmActive := CONTROLLER_DIAGNOSTICS.Status.dwModuleAlarm;
astAlarmSource[22].xGlobalError := TRUE;

ALARM_MANAGER(
    xControllerWarningResetAllowed := NOT CONTROLLER_DIAGNOSTICS.Status.xMemoryWarning
        OR CONTROLLER_DIAGNOSTICS.Status.xWarningResetAllowed,
	xResetWarnings := GVL_ALARM.Command.xResetWarnings,
	astAdditionalCellWarning := astAdditionalCellWarning,
	Sources := astAlarmSource,
	Status => GVL_ALARM.Status
);
IF ALARM_MANAGER.xEventsUpdated OR NOT xHmiTablesInitialized THEN
    GVL_ALARM.Events := ALARM_MANAGER.Events;
END_IF;

(* ---- PLC_PRG.RunCellControl.st ---- *)
METHOD PRIVATE RunCellControl

// --- BEGIN IMPLEMENTATION ---

// Выключенные станки, магазины и ГК не требуют настройки своих точек.
// Общая безопасная точка обязательна при любом составе автоцикла.
xCellPointsReady := GVL_POINT.Points[E_POINT_NAME.HOME_SAFETY].xConfigured;
FOR uiMachine := UINT#1 TO UINT#3 DO
	IF GVL_MACHINE.Status[uiMachine].xEnabled THEN
		xCellPointsReady := xCellPointsReady AND axMachinePointsReady[uiMachine];
	END_IF;
END_FOR;
FOR uiMagazine := UINT#1 TO UINT#2 DO
	IF GVL_MAGAZINE.astStatus[uiMagazine].xEnabled THEN
		xCellPointsReady := xCellPointsReady AND axMagazinePointsReady[uiMagazine];
	END_IF;
	IF GVL_GEOMETRY_CONTROL.astStatus[uiMagazine].xEnabled THEN
		xCellPointsReady := xCellPointsReady
			AND GVL_GEOMETRY_CONTROL.astStatus[uiMagazine].xConfigured;
	END_IF;
END_FOR;

uiMagazine := GVL_CELL_MANAGER.Status.uiActiveMagazine;
IF (uiMagazine < UINT#1) OR (uiMagazine > UINT#2) THEN
	uiMagazine := UINT#1;
END_IF;

TYPE_CONFIG(
	xTestInitialize := xTestInitializePulse,
	stTestScenario := GVL_HMI.stTestScenario,
	Command := GVL_HMI.stMultiType.Command,
	xCellRunning := GVL_CELL_MANAGER.Status.xRunning,
	xMotionBusy := xMotionBusy,
	stRobotStatus := GVL_ROBOT.Status,
	astMagazineStatus := GVL_MAGAZINE.astStatus,
	astMachineStatus := GVL_MACHINE.Status,
	uiRows := GVL_CELL_SETTINGS.MagazineRows,
	uiColumns := GVL_CELL_SETTINGS.MagazineColumns,
	Config => GVL_MULTI_TYPE.Config,
	Status => GVL_MULTI_TYPE.ConfigStatus
);

CELL_MANAGER(
	axMagazineAutoSwapPending := axTwinAutoSwapPending,
	axMagazineExchangeInProgress := axTwinMagazineExchangeInProgress,
	xMagazineExchangeActive := (GVL_TWO_PALLET.uiMode = 1) AND (
		GVL_TWO_PALLET.astStatus[1].xBusy OR GVL_TWO_PALLET.astStatus[2].xBusy
		OR GVL_TWO_PALLET.astStatus[1].xCompleted OR GVL_TWO_PALLET.astStatus[2].xCompleted),
	xStart := GVL_CELL_CONTROL.xStart,
	xStop := GVL_CELL_CONTROL.xStop,
	xTestAbort := xTestAbortActive,
	xResetRequest := GVL_HMI.xCellReset,
	xReset := GVL_CELL_CONTROL.xReset,
	xOperatorChoice := GVL_HMI.xCellOperatorChoice,
	xOperatorCancel := GVL_HMI.xCellOperatorCancel,
	uiOperatorChoice := GVL_HMI.uiCellOperatorChoice,
	xManual := GVL_CELL_CONTROL.xManual,
	xIoManual := xIoManualActive,
	uiModeRejectReason := uiCellModeRejectReason,
	xSettingsRejected := xCellSettingRejected,
	xIoOverrideRejected := xIoOverrideRejected,
    xIoDoRejected := xIoDoRejected,
    xIoEmergencyResetRejected := xIoEmergencyResetRejected,
    xIoEmergencyStopActive := GVL_HMI.xIoEmergencyStopActive,
	xGlobalError := GVL_CELL_CONTROL.xGlobalError,
	xSafetyReady := CELL_SAFETY.Status.xReady AND NOT CONTROLLER_DIAGNOSTICS.Status.xAlarmActive,
	xDrivesReady := xDrivesReady,
	xMotionBusy := xMotionBusy,
	xRobotInterfaceReady := xRobotInterfaceReady,
	lrRobotActualX := lrRobotActualX,
	lrRobotActualY := lrRobotActualY,
	lrRobotActualZ := lrRobotActualZ,
	stSafetyHomePoint := GVL_POINT.Points[E_POINT_NAME.HOME_SAFETY],
	lrSafetyHomeToleranceX := GVL_CELL_SETTINGS.lrSafetyHomeToleranceX,
	lrSafetyHomeToleranceY := GVL_CELL_SETTINGS.lrSafetyHomeToleranceY,
	lrSafetyHomeToleranceZ := GVL_CELL_SETTINGS.lrSafetyHomeToleranceZ,
	lrStoppedPoseTolerance := GVL_CELL_SETTINGS.lrStoppedPoseTolerance,
	Config := GVL_MULTI_TYPE.Config,
	xConfigurationValid := GVL_MULTI_TYPE.ConfigStatus.xConfigurationValid,
	xPointsConfigured := xCellPointsReady,
	stRobotStatus := GVL_ROBOT.Status,
	astMagazineStatus := GVL_MAGAZINE.astStatus,
	astMachineStatus := GVL_MACHINE.Status,
	astMachineDiag := GVL_MACHINE.Diag,
	FaultRequest := stCellFaultRequest,
	Command => GVL_CELL_MANAGER.Command,
	Status => GVL_CELL_MANAGER.Status,
	Diag => GVL_CELL_MANAGER.Diag,
	Error => GVL_CELL_MANAGER.Error,
	CycleStatus => GVL_MULTI_TYPE.CycleStatus
);

// Сначала снимаем команды обоих владельцев, затем маршрутизируем единственную
// команду менеджера выбранному магазину.
// Общий Disable ячейки не отключает независимо включённые магазины.
FOR uiMagazine := UINT#1 TO UINT#2 DO
	GVL_MAGAZINE.astAutoCommand[uiMagazine].xEnable := FALSE;
	GVL_MAGAZINE.astAutoCommand[uiMagazine].xDisable := FALSE;
	GVL_MAGAZINE.astAutoCommand[uiMagazine].xExecute := FALSE;
	GVL_MAGAZINE.astAutoCommand[uiMagazine].xStop := FALSE;
	GVL_MAGAZINE.astAutoCommand[uiMagazine].eOperation := E_MAGAZINE_OPERATION.NONE;
	GVL_MAGAZINE.astAutoCommand[uiMagazine].iTakeSlot := SINT#0;
	GVL_MAGAZINE.astAutoCommand[uiMagazine].iPutSlot := SINT#0;
END_FOR;
IF (GVL_CELL_MANAGER.Status.uiActiveMagazine >= UINT#1)
AND (GVL_CELL_MANAGER.Status.uiActiveMagazine <= UINT#2) THEN
	GVL_MAGAZINE.astAutoCommand[GVL_CELL_MANAGER.Status.uiActiveMagazine] :=
		GVL_CELL_MANAGER.Command.stMagazine;
	GVL_MAGAZINE.astAutoCommand[GVL_CELL_MANAGER.Status.uiActiveMagazine].xEnable := FALSE;
END_IF;

(* ---- PLC_PRG.RunGeometryControl.st ---- *)
METHOD PRIVATE RunGeometryControl

// --- BEGIN IMPLEMENTATION ---

xGeometryEnvironmentChanged := NOT xGeometryInitialized
	OR (eGeometryPreviousEnvironment <> GVL_CELL_SETTINGS.eTestEnvironment);
GVL_GEOMETRY_CONTROL.uiEnvironment := TO_UINT(GVL_CELL_SETTINGS.eTestEnvironment);
GVL_GEOMETRY_CONTROL.xSupported := NOT GVL_HMI.xModbusMode
	AND (GVL_CELL_SETTINGS.eTestEnvironment <> E_CELL_TEST_ENVIRONMENT.SC500_BENCH);
IF xGeometryEnvironmentChanged THEN
	FOR uiGeometry := UINT#1 TO UINT#2 DO
		IF GVL_CELL_SETTINGS.eTestEnvironment = E_CELL_TEST_ENVIRONMENT.NORMAL THEN
			GVL_GEOMETRY_CONTROL.astActiveMemory[uiGeometry] := Persistent_Value.astMemory[uiGeometry];
		ELSE GVL_GEOMETRY_CONTROL.astActiveMemory[uiGeometry] := GVL_GEOMETRY_CONTROL.astSimulationMemory[uiGeometry]; END_IF;
		GVL_GEOMETRY_CONTROL.astSignals[uiGeometry].xReserve := FALSE;
		GVL_GEOMETRY_CONTROL.astSignals[uiGeometry].xDeposited := FALSE;
		GVL_GEOMETRY_CONTROL.astSignals[uiGeometry].xReleased := FALSE;
		GVL_GEOMETRY_CONTROL.astSignals[uiGeometry].xRobotInteraction := FALSE;
	END_FOR;
	FOR uiGeometryMachine := UINT#1 TO UINT#3 DO
		IF GVL_CELL_SETTINGS.eTestEnvironment = E_CELL_TEST_ENVIRONMENT.NORMAL THEN
			GVL_GEOMETRY_CONTROL.astCalls[uiGeometryMachine] := Persistent_Value.astRetainCalls[uiGeometryMachine];
			GVL_GEOMETRY_CONTROL.auiActiveCount[uiGeometryMachine] := Persistent_Value.auiCount[uiGeometryMachine];
		ELSE
			GVL_GEOMETRY_CONTROL.astCalls[uiGeometryMachine] := GVL_GEOMETRY_CONTROL.astSimulationCalls[uiGeometryMachine];
			GVL_GEOMETRY_CONTROL.auiActiveCount[uiGeometryMachine] := GVL_GEOMETRY_CONTROL.auiSimulationCount[uiGeometryMachine];
		END_IF;
		IF (GVL_GEOMETRY_CONTROL.astCalls[uiGeometryMachine].uiState = UINT#2)
		OR (GVL_GEOMETRY_CONTROL.astCalls[uiGeometryMachine].uiState = UINT#3) THEN
			GVL_GEOMETRY_CONTROL.astCalls[uiGeometryMachine].uiState := UINT#7;
			GVL_GEOMETRY_CONTROL.astCalls[uiGeometryMachine].uiReason := UINT#5;
			F_GEOMETRY_EVENT(Call := GVL_GEOMETRY_CONTROL.astCalls[uiGeometryMachine]);
		END_IF;
	END_FOR;
	xGeometryInitialized := TRUE;
	eGeometryPreviousEnvironment := GVL_CELL_SETTINGS.eTestEnvironment;
END_IF;
// Only the accepted simulation buffer can reset virtual station inventory.
IF xTestInitializePulse AND (GVL_CELL_SETTINGS.eTestEnvironment = E_CELL_TEST_ENVIRONMENT.SIMULATION) THEN
	FOR uiGeometry := UINT#1 TO UINT#2 DO
		udiTestGeometryProduced := GVL_GEOMETRY_CONTROL.astActiveMemory[uiGeometry].udiProducedPartsTotal;
		GVL_GEOMETRY_CONTROL.astActiveMemory[uiGeometry] := stTestEmptyGeometryMemory;
		GVL_GEOMETRY_CONTROL.astActiveMemory[uiGeometry].udiProducedPartsTotal := udiTestGeometryProduced;
		GVL_GEOMETRY_CONTROL.astSimulationMemory[uiGeometry] := GVL_GEOMETRY_CONTROL.astActiveMemory[uiGeometry];
		GVL_GEOMETRY_CONTROL.astSignals[uiGeometry].xReserve := FALSE;
		GVL_GEOMETRY_CONTROL.astSignals[uiGeometry].xDeposited := FALSE;
		GVL_GEOMETRY_CONTROL.astSignals[uiGeometry].xReleased := FALSE;
		GVL_GEOMETRY_CONTROL.astSignals[uiGeometry].xRobotInteraction := FALSE;
		GVL_GEOMETRY_CONTROL.axSimulationAlarm[uiGeometry] := FALSE;
	END_FOR;
	FOR uiGeometryMachine := UINT#1 TO UINT#3 DO
		GVL_GEOMETRY_CONTROL.astCalls[uiGeometryMachine] := stTestEmptyGeometryCall;
		GVL_GEOMETRY_CONTROL.auiActiveCount[uiGeometryMachine] := UINT#0;
		IF GVL_HMI.stTestScenario.axGeometryCall[uiGeometryMachine] THEN
			Persistent_Value.udiNextCallId := Persistent_Value.udiNextCallId + UDINT#1;
			IF Persistent_Value.udiNextCallId = UDINT#0 THEN Persistent_Value.udiNextCallId := UDINT#1; END_IF;
			GVL_GEOMETRY_CONTROL.astCalls[uiGeometryMachine].udiId := Persistent_Value.udiNextCallId;
			GVL_GEOMETRY_CONTROL.astCalls[uiGeometryMachine].uiMachine := uiGeometryMachine;
			GVL_GEOMETRY_CONTROL.astCalls[uiGeometryMachine].uiProductType := GVL_HMI.stTestScenario.auiMachineType[uiGeometryMachine];
			GVL_GEOMETRY_CONTROL.astCalls[uiGeometryMachine].uiState := UINT#1;
			GVL_GEOMETRY_CONTROL.astCalls[uiGeometryMachine].xForced := TRUE;
		END_IF;
	END_FOR;
END_IF;
FOR uiGeometry := UINT#1 TO UINT#2 DO
	GVL_GEOMETRY_CONTROL.auiAction[uiGeometry] := UINT#0;
	IF GVL_CELL_SETTINGS.eTestEnvironment = E_CELL_TEST_ENVIRONMENT.NORMAL THEN
		GVL_GEOMETRY_CONTROL.astActiveConfig[uiGeometry] := Persistent_Value.astConfig[uiGeometry];
	ELSE GVL_GEOMETRY_CONTROL.astActiveConfig[uiGeometry] := Persistent_Value.astSimulationConfig[uiGeometry]; END_IF;
END_FOR;
GVL_GEOMETRY_CONTROL.xAutoChangeAllowed := GVL_GEOMETRY_CONTROL.xSupported
	AND xHmiConnectionAlive AND NOT GVL_HMI.xTestSessionActive AND NOT GVL_CELL_CONTROL.xGlobalError;
GVL_GEOMETRY_CONTROL.xSettingsAllowed := GVL_GEOMETRY_CONTROL.xSupported
	AND GVL_CELL_SETTINGS.xCellSettingsChangeAllowed AND xHmiConnectionAlive
	AND NOT GVL_GEOMETRY_CONTROL.astStatus[1].xDriveRunning AND NOT GVL_GEOMETRY_CONTROL.astStatus[2].xDriveRunning
	AND NOT GVL_GEOMETRY_CONTROL.astStatus[1].xResetBusy AND NOT GVL_GEOMETRY_CONTROL.astStatus[2].xResetBusy
	AND NOT GVL_GEOMETRY_CONTROL.astStatus[1].xReserved AND NOT GVL_GEOMETRY_CONTROL.astStatus[2].xReserved
	AND NOT GVL_GEOMETRY_CONTROL.astSignals[1].xRobotInteraction AND NOT GVL_GEOMETRY_CONTROL.astSignals[2].xRobotInteraction
	AND NOT GEOMETRY[1].xRunOutput AND NOT GEOMETRY[2].xRunOutput;
FOR uiGeometryMachine := UINT#1 TO UINT#3 DO
	GVL_GEOMETRY_CONTROL.axCallAllowed[uiGeometryMachine] := GVL_GEOMETRY_CONTROL.xAutoChangeAllowed
		AND GVL_MACHINE.Status[uiGeometryMachine].xEnabled
		AND ((GVL_GEOMETRY_CONTROL.astCalls[uiGeometryMachine].uiState <= UINT#1)
			OR (GVL_GEOMETRY_CONTROL.astCalls[uiGeometryMachine].uiState > UINT#3))
		AND (GVL_GEOMETRY_CONTROL.astStatus[1].xEnabled OR GVL_GEOMETRY_CONTROL.astStatus[2].xEnabled);
	GVL_GEOMETRY_CONTROL.axCancelAllowed[uiGeometryMachine] := GVL_GEOMETRY_CONTROL.xAutoChangeAllowed
		AND (GVL_GEOMETRY_CONTROL.astCalls[uiGeometryMachine].uiState = UINT#1);
END_FOR;

// Упакованный канал: подготовка payload -> CommandSeq -> Result -> Ack.
udiGeometryRequest := GVL_HMI.udiGeometryCommandSeq;
xGeometryRequestFresh := FALSE;
IF (udiGeometryRequest <> UDINT#0) AND (udiGeometryRequest <> GVL_HMI.udiGeometryAckSeq) THEN
	stGeometryRequest := GVL_HMI.stGeometryRequest;
	GVL_HMI.uiGeometryResult := UINT#2;
	IF NOT IsHmiCommandFresh(udiIssuedAtMs := GVL_HMI.udiGeometryIssuedAtMs) THEN
		GVL_HMI.uiGeometryResult := UINT#4;
	ELSIF xHmiConnectionAlive THEN
		xGeometryRequestFresh := TRUE;
		IF (stGeometryRequest.uiAction = UINT#8) AND (stGeometryRequest.uiMachine >= UINT#1)
		AND (stGeometryRequest.uiMachine <= UINT#3) THEN
			uiGeometryMachine := stGeometryRequest.uiMachine;
			IF GVL_GEOMETRY_CONTROL.axCallAllowed[uiGeometryMachine] THEN
				IF GVL_GEOMETRY_CONTROL.astCalls[uiGeometryMachine].uiState = UINT#1 THEN
					stGeometryCall := GVL_GEOMETRY_CONTROL.astCalls[uiGeometryMachine];
				ELSE
					Persistent_Value.udiNextCallId := Persistent_Value.udiNextCallId + UDINT#1;
					IF Persistent_Value.udiNextCallId = UDINT#0 THEN Persistent_Value.udiNextCallId := UDINT#1; END_IF;
					stGeometryCall := stGeometryEmptyCall;
					stGeometryCall.udiId := Persistent_Value.udiNextCallId;
					stGeometryCall.uiMachine := uiGeometryMachine;
					stGeometryCall.uiProductType := GVL_MULTI_TYPE.Config.auiMachineType[uiGeometryMachine];
				END_IF;
				stGeometryCall.xForced := TRUE; stGeometryCall.uiState := UINT#1;
				GVL_GEOMETRY_CONTROL.astCalls[uiGeometryMachine] := stGeometryCall;
				GVL_GEOMETRY_CONTROL.auiActiveCount[uiGeometryMachine] := UINT#0;
				F_GEOMETRY_EVENT(Call := stGeometryCall); GVL_HMI.uiGeometryResult := UINT#1;
			END_IF;
		ELSIF (stGeometryRequest.uiAction = UINT#12) AND (stGeometryRequest.uiMachine >= UINT#1)
		AND (stGeometryRequest.uiMachine <= UINT#3) THEN
			uiGeometryMachine := stGeometryRequest.uiMachine;
			IF GVL_GEOMETRY_CONTROL.axCancelAllowed[uiGeometryMachine] THEN
				GVL_GEOMETRY_CONTROL.astCalls[uiGeometryMachine].uiState := UINT#6;
				F_GEOMETRY_EVENT(Call := GVL_GEOMETRY_CONTROL.astCalls[uiGeometryMachine]); GVL_HMI.uiGeometryResult := UINT#1;
			END_IF;
		ELSIF (stGeometryRequest.uiAction = UINT#9) AND GVL_GEOMETRY_CONTROL.xAutoChangeAllowed
		AND (stGeometryRequest.udiValue <= UDINT#1) THEN
			Persistent_Value.xAutoEnabled := stGeometryRequest.udiValue = UDINT#1;
			GVL_HMI.uiGeometryResult := UINT#1;
		ELSIF (stGeometryRequest.uiAction = UINT#10) AND GVL_GEOMETRY_CONTROL.xAutoChangeAllowed
		AND (stGeometryRequest.uiMachine <= UINT#3) AND (stGeometryRequest.udiValue >= UDINT#1)
		AND (stGeometryRequest.udiValue <= UDINT#10000) THEN
			FOR uiGeometryMachine := UINT#1 TO UINT#3 DO
				IF (stGeometryRequest.uiMachine = UINT#0) OR (stGeometryRequest.uiMachine = uiGeometryMachine) THEN
					Persistent_Value.auiPeriod[uiGeometryMachine] := UDINT_TO_UINT(stGeometryRequest.udiValue);
				END_IF;
			END_FOR;
			GVL_HMI.uiGeometryResult := UINT#1;
		ELSIF (stGeometryRequest.uiAction = UINT#16) AND GVL_GEOMETRY_CONTROL.xSettingsAllowed THEN
			CASE stGeometryRequest.uiMachine OF
				UINT#1: IF stGeometryRequest.udiValue <= UDINT#1 THEN Persistent_Value.xWaitWhenOccupied := stGeometryRequest.udiValue = UDINT#1; GVL_HMI.uiGeometryResult := UINT#1; END_IF;
				UINT#2: IF (stGeometryRequest.udiValue >= UDINT#100) AND (stGeometryRequest.udiValue <= UDINT#600000) THEN Persistent_Value.tTransportTimeout := UDINT_TO_TIME(stGeometryRequest.udiValue); GVL_HMI.uiGeometryResult := UINT#1; END_IF;
				UINT#3: IF (stGeometryRequest.udiValue >= UDINT#100) AND (stGeometryRequest.udiValue <= UDINT#60000) THEN Persistent_Value.tDriveFeedbackTimeout := UDINT_TO_TIME(stGeometryRequest.udiValue); GVL_HMI.uiGeometryResult := UINT#1; END_IF;
				UINT#4: IF (stGeometryRequest.udiValue >= UDINT#100) AND (stGeometryRequest.udiValue <= UDINT#10000) THEN Persistent_Value.tResetPulse := UDINT_TO_TIME(stGeometryRequest.udiValue); GVL_HMI.uiGeometryResult := UINT#1; END_IF;
				UINT#5: IF (stGeometryRequest.udiValue >= UDINT#1000) AND (stGeometryRequest.udiValue <= UDINT#3600000) THEN Persistent_Value.tWaitWarningTimeout := UDINT_TO_TIME(stGeometryRequest.udiValue); GVL_HMI.uiGeometryResult := UINT#1; END_IF;
			END_CASE;
		ELSIF (stGeometryRequest.uiStation >= UINT#1) AND (stGeometryRequest.uiStation <= UINT#2) THEN
			uiGeometry := stGeometryRequest.uiStation;
			IF (stGeometryRequest.uiAction >= UINT#1) AND (stGeometryRequest.uiAction <= UINT#7) THEN
				GVL_GEOMETRY_CONTROL.auiAction[uiGeometry] := stGeometryRequest.uiAction;
			ELSIF (stGeometryRequest.uiAction = UINT#11) AND GVL_GEOMETRY_CONTROL.xSupported
			AND GVL_POINT_MANAGER.PointManager.Diag.xXLimitValid
			AND GVL_POINT_MANAGER.PointManager.Diag.xYLimitValid
			AND GVL_POINT_MANAGER.PointManager.Diag.xZLimitValid THEN
				stGeometryConfig := stGeometryRequest.Config;
				stGeometryConfig.lrChangeZ := stGeometryConfig.lrSafeZ;
				xGeometryConfigValid := (stGeometryConfig.lrSpeedFactor >= 0.1) AND (stGeometryConfig.lrSpeedFactor <= 1.0)
					AND (stGeometryConfig.lrSafeZ < 0.0) AND (stGeometryConfig.lrSafeZ >= -10000.0)
					AND (stGeometryConfig.lrX >= GVL_POINT_MANAGER.PointManager.Diag.lrX_MinLimit)
					AND (stGeometryConfig.lrX <= GVL_POINT_MANAGER.PointManager.Diag.lrX_MaxLimit)
					AND (stGeometryConfig.lrY >= GVL_POINT_MANAGER.PointManager.Diag.lrY_MinLimit)
					AND (stGeometryConfig.lrY <= GVL_POINT_MANAGER.PointManager.Diag.lrY_MaxLimit)
					AND (stGeometryConfig.lrZ >= GVL_POINT_MANAGER.PointManager.Diag.lrZ_MinLimit)
					AND (stGeometryConfig.lrZ <= GVL_POINT_MANAGER.PointManager.Diag.lrZ_MaxLimit)
					AND ((stGeometryConfig.lrZ + stGeometryConfig.lrSafeZ) >= GVL_POINT_MANAGER.PointManager.Diag.lrZ_MinLimit);
				IF xGeometryConfigValid THEN
					stGeometryConfig.xConfigured := TRUE;
					IF GVL_CELL_SETTINGS.eTestEnvironment = E_CELL_TEST_ENVIRONMENT.NORMAL THEN Persistent_Value.astConfig[uiGeometry] := stGeometryConfig;
					ELSE Persistent_Value.astSimulationConfig[uiGeometry] := stGeometryConfig; END_IF;
					GVL_GEOMETRY_CONTROL.astActiveConfig[uiGeometry] := stGeometryConfig; GVL_HMI.uiGeometryResult := UINT#1;
				END_IF;
			ELSIF (stGeometryRequest.uiAction = UINT#13) AND GVL_GEOMETRY_CONTROL.astStatus[uiGeometry].xPointWriteAllowed
			AND GVL_HMI.xPointEditorCaptureAllowed THEN
				GVL_HMI.stGeometryCapture := GVL_GEOMETRY_CONTROL.astActiveConfig[uiGeometry];
				GVL_HMI.stGeometryCapture.lrX := lrRobotActualX; GVL_HMI.stGeometryCapture.lrY := lrRobotActualY;
				GVL_HMI.stGeometryCapture.lrZ := lrRobotActualZ; GVL_HMI.uiGeometryResult := UINT#1;
			ELSIF ((stGeometryRequest.uiAction = UINT#14) OR (stGeometryRequest.uiAction = UINT#15))
			AND GVL_CELL_SETTINGS.xErrorSimulationEnabled
			AND (GVL_CELL_SETTINGS.eTestEnvironment = E_CELL_TEST_ENVIRONMENT.SIMULATION)
			AND GVL_GEOMETRY_CONTROL.xSupported THEN
				GVL_GEOMETRY_CONTROL.axSimulationAlarm[uiGeometry] := stGeometryRequest.uiAction = UINT#14;
				GVL_HMI.uiGeometryResult := UINT#1;
			END_IF;
		END_IF;
	END_IF;
END_IF;

FOR uiGeometry := UINT#1 TO UINT#2 DO
	xGeometryStopAttempt := FALSE;
	IF (GVL_HMI.audiGeometryStopSeq[uiGeometry] <> UDINT#0)
	AND (GVL_HMI.audiGeometryStopSeq[uiGeometry] <> GVL_HMI.audiGeometryStopAck[uiGeometry]) THEN
		GVL_GEOMETRY_CONTROL.auiAction[uiGeometry] := UINT#6;
		xGeometryStopAttempt := TRUE;
		GVL_HMI.audiGeometryStopAck[uiGeometry] := GVL_HMI.audiGeometryStopSeq[uiGeometry];
	END_IF;
	IF GVL_CELL_SETTINGS.eTestEnvironment <> E_CELL_TEST_ENVIRONMENT.NORMAL THEN
		GEOMETRY_SIM[uiGeometry](xInitialize := xGeometryEnvironmentChanged OR xTestInitializePulse,
			xRun := GEOMETRY[uiGeometry].xRunOutput, xReset := GEOMETRY[uiGeometry].xResetOutput,
			xDeposited := GVL_GEOMETRY_CONTROL.astSignals[uiGeometry].xDeposited,
			udiPartId := GVL_GEOMETRY_CONTROL.astSignals[uiGeometry].Call.udiId,
			xRemove := GEOMETRY[uiGeometry].xSimulationEmptyConfirmed,
			xAlarm := GVL_GEOMETRY_CONTROL.axSimulationAlarm[uiGeometry],
			uiTimeFactor := SEL(GVL_CELL_SETTINGS.xSimulationAccelerationActive, UINT#1, GVL_CELL_SETTINGS.uiSimulationTimeFactorApplied));
		xGeometryDriveAlarm := GEOMETRY_SIM[uiGeometry].xDriveAlarm;
		xGeometryDriveRunning := GEOMETRY_SIM[uiGeometry].xDriveRunning;
		xGeometryPartAtEnd := GEOMETRY_SIM[uiGeometry].xPartAtEnd;
	ELSE
		uiGeometryDi := UINT#81 + (uiGeometry - UINT#1) * UINT#2;
		xGeometryDriveAlarm := xPhysicalNormal AND (GVL_PHYSICAL_IO.xMappingVerified OR axIoForced[uiGeometryDi]) AND axPhysicalRaw[uiGeometryDi];
		xGeometryDriveRunning := xPhysicalNormal AND (GVL_PHYSICAL_IO.xMappingVerified OR axIoForced[uiGeometryDi + UINT#1]) AND axPhysicalRaw[uiGeometryDi + UINT#1];
		xGeometryPartAtEnd := GVL_PHYSICAL_IO.axGkPartAtEnd[uiGeometry];
	END_IF;
	stGeometrySignals := GVL_GEOMETRY_CONTROL.astSignals[uiGeometry];
	// Ручное движение также считается работой с ГК; состояние последней точки
	// удерживает блокировку ленты вплоть до подтверждённого отхода.
	IF uiGeometry = UINT#1 THEN
		stGeometrySignals.xRobotInteraction := stGeometrySignals.xRobotInteraction
			OR (GVL_ROBOT.Status.eCurrentPoint = E_POINT_NAME.GEOMETRY_1_PLACE)
			OR (GVL_ROBOT.Status.eCurrentPoint = E_POINT_NAME.GEOMETRY_1_CHANGE)
			OR (GVL_ROBOT.Status.xBusy AND ((GVL_ROBOT.Command.eSetPoint = E_POINT_NAME.GEOMETRY_1_PLACE)
				OR (GVL_ROBOT.Command.eSetPoint = E_POINT_NAME.GEOMETRY_1_CHANGE)));
	ELSE
		stGeometrySignals.xRobotInteraction := stGeometrySignals.xRobotInteraction
			OR (GVL_ROBOT.Status.eCurrentPoint = E_POINT_NAME.GEOMETRY_2_PLACE)
			OR (GVL_ROBOT.Status.eCurrentPoint = E_POINT_NAME.GEOMETRY_2_CHANGE)
			OR (GVL_ROBOT.Status.xBusy AND ((GVL_ROBOT.Command.eSetPoint = E_POINT_NAME.GEOMETRY_2_PLACE)
				OR (GVL_ROBOT.Command.eSetPoint = E_POINT_NAME.GEOMETRY_2_CHANGE)));
	END_IF;
	GEOMETRY[uiGeometry](xInitialize := xGeometryEnvironmentChanged OR xTestInitializePulse, uiAction := GVL_GEOMETRY_CONTROL.auiAction[uiGeometry],
		xSupported := GVL_GEOMETRY_CONTROL.xSupported AND ((GVL_CELL_SETTINGS.eTestEnvironment <> E_CELL_TEST_ENVIRONMENT.NORMAL) OR GVL_PHYSICAL_IO.xMappingVerified),
		xSimulation := GVL_CELL_SETTINGS.eTestEnvironment <> E_CELL_TEST_ENVIRONMENT.NORMAL,
		xGlobalError := GVL_CELL_CONTROL.xGlobalError, xManual := GVL_CELL_CONTROL.xManual,
		xCellRunning := GVL_CELL_MANAGER.Status.xRunning, xRobotBusy := GVL_ROBOT.Status.xBusy,
		xMotionBusy := xMotionBusy, xHmiAlive := xHmiConnectionAlive, xIoManual := xIoManualActive,
		xReset := GVL_CELL_CONTROL.xReset, xDriveAlarm := xGeometryDriveAlarm,
		xDriveRunning := xGeometryDriveRunning, xPartAtEnd := xGeometryPartAtEnd,
		rSimulationTravel := GEOMETRY_SIM[uiGeometry].rTravel,
		Signals := stGeometrySignals, Config := GVL_GEOMETRY_CONTROL.astActiveConfig[uiGeometry],
		tTransport := Persistent_Value.tTransportTimeout, tFeedback := Persistent_Value.tDriveFeedbackTimeout,
		tResetPulse := Persistent_Value.tResetPulse,
		uiTimeFactor := SEL(GVL_CELL_SETTINGS.xSimulationAccelerationActive, UINT#1, GVL_CELL_SETTINGS.uiSimulationTimeFactorApplied),
		Memory := GVL_GEOMETRY_CONTROL.astActiveMemory[uiGeometry], Status => GVL_GEOMETRY_CONTROL.astStatus[uiGeometry],
		Warning => GVL_GEOMETRY_CONTROL.astWarning[uiGeometry]);
	GVL_GEOMETRY_CONTROL.astStatus[uiGeometry].xConfigAllowed := GVL_GEOMETRY_CONTROL.astStatus[uiGeometry].xConfigAllowed AND GVL_HMI.xPointEditorSaveAllowed;
	// Только доступность канала данных и лимитов; физическая карта, Home,
	// режим, ошибки, движение и состояние станции не ограничивают SAVE.
	GVL_GEOMETRY_CONTROL.astStatus[uiGeometry].xPointWriteAllowed := GVL_GEOMETRY_CONTROL.xSupported
		AND xHmiConnectionAlive AND GVL_POINT_MANAGER.PointManager.Diag.xXLimitValid
		AND GVL_POINT_MANAGER.PointManager.Diag.xYLimitValid
		AND GVL_POINT_MANAGER.PointManager.Diag.xZLimitValid;
	GVL_GEOMETRY_CONTROL.astStatus[uiGeometry].xSimulationAlarmAllowed := GVL_GEOMETRY_CONTROL.xSupported
		AND (GVL_CELL_SETTINGS.eTestEnvironment = E_CELL_TEST_ENVIRONMENT.SIMULATION)
		AND GVL_CELL_SETTINGS.xErrorSimulationEnabled AND xHmiConnectionAlive;
	IF xGeometryRequestFresh AND NOT xGeometryStopAttempt
	AND (udiGeometryRequest <> UDINT#0) AND (udiGeometryRequest <> GVL_HMI.udiGeometryAckSeq)
	AND (stGeometryRequest.uiStation = uiGeometry) AND (stGeometryRequest.uiAction >= UINT#1) AND (stGeometryRequest.uiAction <= UINT#7) THEN
		IF GEOMETRY[uiGeometry].xCommandAccepted THEN GVL_HMI.uiGeometryResult := UINT#1; END_IF;
	END_IF;
	// Точки ГК независимы от механики/баз палет и от включения магазина.
	IF uiGeometry = UINT#1 THEN eGeometryPlace := E_POINT_NAME.GEOMETRY_1_PLACE; eGeometrySafe := E_POINT_NAME.GEOMETRY_1_SAFE; eGeometryChange := E_POINT_NAME.GEOMETRY_1_CHANGE;
	ELSE eGeometryPlace := E_POINT_NAME.GEOMETRY_2_PLACE; eGeometrySafe := E_POINT_NAME.GEOMETRY_2_SAFE; eGeometryChange := E_POINT_NAME.GEOMETRY_2_CHANGE; END_IF;
	GVL_POINT.Points[eGeometryPlace].X := GVL_GEOMETRY_CONTROL.astActiveConfig[uiGeometry].lrX;
	GVL_POINT.Points[eGeometryPlace].Y := GVL_GEOMETRY_CONTROL.astActiveConfig[uiGeometry].lrY;
	GVL_POINT.Points[eGeometryPlace].Z := GVL_GEOMETRY_CONTROL.astActiveConfig[uiGeometry].lrZ;
	GVL_POINT.Points[eGeometryPlace].MagazineSafeZ := GVL_GEOMETRY_CONTROL.astActiveConfig[uiGeometry].lrSafeZ;
	GVL_POINT.Points[eGeometryPlace].MagazineChangeZ := LREAL#0.0;
	GVL_POINT.Points[eGeometryPlace].SpeedFactor := GVL_GEOMETRY_CONTROL.astActiveConfig[uiGeometry].lrSpeedFactor;
	GVL_POINT.Points[eGeometryPlace].xConfigured := GVL_GEOMETRY_CONTROL.astActiveConfig[uiGeometry].xConfigured;
	GVL_POINT.Points[eGeometrySafe] := GVL_POINT.Points[eGeometryPlace];
	GVL_POINT.Points[eGeometrySafe].Z := GVL_POINT.Points[eGeometryPlace].Z + GVL_GEOMETRY_CONTROL.astActiveConfig[uiGeometry].lrSafeZ;
	GVL_POINT.Points[eGeometryChange] := GVL_POINT.Points[eGeometrySafe]; // Legacy CHANGE совпадает с SAFE_Z
END_FOR;
IF (udiGeometryRequest <> UDINT#0) AND (udiGeometryRequest <> GVL_HMI.udiGeometryAckSeq) THEN
	IF GVL_HMI.uiGeometryResult <> UINT#1 THEN
		GVL_GEOMETRY_CONTROL.stCellWarning.uiCode := UINT#51;
		GVL_GEOMETRY_CONTROL.stCellWarning.udiSequence := GVL_GEOMETRY_CONTROL.stCellWarning.udiSequence + UDINT#1;
	END_IF;
	GVL_HMI.udiGeometryAckSeq := udiGeometryRequest;
END_IF;

(* ---- PLC_PRG.RunMachines.st ---- *)
METHOD PRIVATE RunMachines

// --- BEGIN IMPLEMENTATION ---

// Импульсные команды HMI изменяют сохранённое разрешение работы станка.
FOR uiMachine := 1 TO 3 DO
	IF GVL_HMI.axMachineDisable[uiMachine] THEN
		GVL_HMI.axMachineUsed[uiMachine] := FALSE;
	ELSIF GVL_HMI.axMachineEnable[uiMachine] AND axMachinePointsReady[uiMachine] THEN
		GVL_HMI.axMachineUsed[uiMachine] := TRUE;
	END_IF;
END_FOR;

MACHINE_1.stPoints.eAbove := E_POINT_NAME.MACHINE_1_ABOVE;
MACHINE_1.stPoints.eChuck := E_POINT_NAME.MACHINE_1_CHUCK_POSITION;
MACHINE_1.stPoints.eChuckApproach := E_POINT_NAME.MACHINE_1_CHUCK_APROACH;
MACHINE_1.stPoints.eInside := E_POINT_NAME.MACHINE_1_INSIDE;
MACHINE_1.stPoints.eNone := E_POINT_NAME.NONE;

// NORMAL получает только физическую обратную связь; обе тестовые среды — модель.
IF GVL_CELL_SETTINGS.eTestEnvironment <> E_CELL_TEST_ENVIRONMENT.NORMAL THEN
// Виртуальные устройства исполняют команду предыдущего цикла. Затем слой
// инъекции формирует обратную связь, которую увидит технологический автомат.
MACHINE_1_SIM(
	xTestInitialize := xTestInitializePulse OR xTestAbortActive,
	uiTestInitialState := GVL_HMI.stTestScenario.auiMachineState[1],
	xSafetyDoorOpen := GVL_CELL_SETTINGS.xErrorSimulationEnabled
		AND GVL_HMI.axMachineSimSafetyDoorOpen[1],
	Command := GVL_MACHINE.Command[1].stIo,
	FaultRequest := astMachineFaultRequest[1],
	xSimulationAccelerationEnable := GVL_CELL_SETTINGS.xSimulationAccelerationActive,
	uiSimulationTimeFactor := GVL_CELL_SETTINGS.uiSimulationTimeFactorApplied,
	tDoorOpenTime := GVL_HMI.tMachineDoorOpenTime,
	tDoorCloseTime := GVL_HMI.tMachineDoorCloseTime,
	tChuckOpenTime := GVL_HMI.tMachineChuckOpenTime,
	tChuckCloseTime := GVL_HMI.tMachineChuckCloseTime,
	tCycleTime := GVL_HMI.tMachineCycleTime[1]
);
MACHINE_2_SIM(
	xTestInitialize := xTestInitializePulse OR xTestAbortActive,
	uiTestInitialState := GVL_HMI.stTestScenario.auiMachineState[2],
	xSafetyDoorOpen := GVL_CELL_SETTINGS.xErrorSimulationEnabled
		AND GVL_HMI.axMachineSimSafetyDoorOpen[2],
	Command := GVL_MACHINE.Command[2].stIo,
	FaultRequest := astMachineFaultRequest[2],
	xSimulationAccelerationEnable := GVL_CELL_SETTINGS.xSimulationAccelerationActive,
	uiSimulationTimeFactor := GVL_CELL_SETTINGS.uiSimulationTimeFactorApplied,
	tDoorOpenTime := GVL_HMI.tMachineDoorOpenTime,
	tDoorCloseTime := GVL_HMI.tMachineDoorCloseTime,
	tChuckOpenTime := GVL_HMI.tMachineChuckOpenTime,
	tChuckCloseTime := GVL_HMI.tMachineChuckCloseTime,
	tCycleTime := GVL_HMI.tMachineCycleTime[2]
);
MACHINE_3_SIM(
	xTestInitialize := xTestInitializePulse OR xTestAbortActive,
	uiTestInitialState := GVL_HMI.stTestScenario.auiMachineState[3],
	xSafetyDoorOpen := GVL_CELL_SETTINGS.xErrorSimulationEnabled
		AND GVL_HMI.axMachineSimSafetyDoorOpen[3],
	Command := GVL_MACHINE.Command[3].stIo,
	FaultRequest := astMachineFaultRequest[3],
	xSimulationAccelerationEnable := GVL_CELL_SETTINGS.xSimulationAccelerationActive,
	uiSimulationTimeFactor := GVL_CELL_SETTINGS.uiSimulationTimeFactorApplied,
	tDoorOpenTime := GVL_HMI.tMachineDoorOpenTime,
	tDoorCloseTime := GVL_HMI.tMachineDoorCloseTime,
	tChuckOpenTime := GVL_HMI.tMachineChuckOpenTime,
	tChuckCloseTime := GVL_HMI.tMachineChuckCloseTime,
	tCycleTime := GVL_HMI.tMachineCycleTime[3]
);

END_IF;
IF GVL_CELL_SETTINGS.eTestEnvironment = E_CELL_TEST_ENVIRONMENT.NORMAL THEN
	astMachineStatusRaw := GVL_MACHINE.astPhysicalInput;
ELSE
	astMachineStatusRaw[1] := MACHINE_1_SIM.Status;
	astMachineStatusRaw[2] := MACHINE_2_SIM.Status;
	astMachineStatusRaw[3] := MACHINE_3_SIM.Status;
END_IF;

MACHINE_1_FAULT(
	xUsePhysicalInput := GVL_CELL_SETTINGS.eTestEnvironment = E_CELL_TEST_ENVIRONMENT.NORMAL,
	Request := astMachineFaultRequest[1],
	MachineStatusRaw := astMachineStatusRaw[1],
	RobotStatusRaw := GVL_ROBOT.Status,
	NominalTimeouts := GVL_CELL_SETTINGS.stMachineTimeouts
);
MACHINE_2_FAULT(
	xUsePhysicalInput := GVL_CELL_SETTINGS.eTestEnvironment = E_CELL_TEST_ENVIRONMENT.NORMAL,
	Request := astMachineFaultRequest[2],
	MachineStatusRaw := astMachineStatusRaw[2],
	RobotStatusRaw := GVL_ROBOT.Status,
	NominalTimeouts := GVL_CELL_SETTINGS.stMachineTimeouts
);
MACHINE_3_FAULT(
	xUsePhysicalInput := GVL_CELL_SETTINGS.eTestEnvironment = E_CELL_TEST_ENVIRONMENT.NORMAL,
	Request := astMachineFaultRequest[3],
	MachineStatusRaw := astMachineStatusRaw[3],
	RobotStatusRaw := GVL_ROBOT.Status,
	NominalTimeouts := GVL_CELL_SETTINGS.stMachineTimeouts
);

MACHINE_1(
	RobotResetRecovery := ROBOT.ResetRecovery,
	xResetCancel := GVL_CELL_CONTROL.xStop OR GVL_CELL_CONTROL.xDisable OR GVL_HMI.xRobotStop,
	xTestInitialize := xTestInitializePulse OR xTestAbortActive,
	uiTestInitialState := GVL_HMI.stTestScenario.auiMachineState[1],
	uiTestProductType := GVL_HMI.stTestScenario.auiMachineType[1],
	xExecute := GVL_CELL_MANAGER.Command.axMachineExecute[1],
	xReset := GVL_HMI.axMachineReset[1],
	xResetGlobal := GVL_CELL_CONTROL.xReset,
	xGlobalError := GVL_CELL_CONTROL.xGlobalError,
	xManualMode := GVL_CELL_CONTROL.xManual,
	xIoManual := xIoManualActive,
	xAutomaticUseEnabled := GVL_HMI.axMachineUsed[1],
	xPointsConfigured := axMachinePointsReady[1],
	xSafetyDoorControlEnabled := GVL_CELL_SETTINGS.eTestEnvironment <> E_CELL_TEST_ENVIRONMENT.NORMAL,
	xHmiOpenSafetyDoor := GVL_HMI.axMachineManualSafetyDoorOpen[1],
	xHmiCloseSafetyDoor := GVL_HMI.axMachineManualSafetyDoorClose[1],
	xHmiOpenHatch := GVL_HMI.axMachineManualHatchOpen[1],
	xHmiCloseHatch := GVL_HMI.axMachineManualHatchClose[1],
	xHmiUnlockHatch := GVL_HMI.axMachineManualHatchUnlock[1],
	xHmiLockHatch := GVL_HMI.axMachineManualHatchLock[1],
	xHmiOpenChuck := GVL_HMI.axMachineManualChuckOpen[1],
	xHmiCloseChuck := GVL_HMI.axMachineManualChuckClose[1],
	xHmiEnable := GVL_HMI.axMachineEnable[1],
	xHmiDisable := GVL_HMI.axMachineDisable[1],
	xHmiSetBlank := GVL_HMI.axMachineSetBlank[1],
	xHmiSetDetail := GVL_HMI.axMachineSetDetail[1],
	xHmiAcceptDoor := GVL_HMI.axMachineAcceptDoor[1],
	xHmiRejectDoor := GVL_HMI.axMachineRejectDoor[1],
	xHmiAcceptRunCNC := GVL_HMI.axMachineAcceptRun[1],
	xHmiRejectRunCNC := GVL_HMI.axMachineRejectRun[1],
	xUseHmiCycleTime := GVL_HMI.xUseHmiCycleTime[1],
	tHmiCycleTime := GVL_HMI.tMachineCycleTime[1],
	stTimeouts := MACHINE_1_FAULT.Timeouts,
	stChangeRecipe := GVL_CELL_SETTINGS.CHANGE_MACHINE,
	stLoadRecipe := GVL_CELL_SETTINGS.LOAD_MACHINE,
	stUnloadRecipe := GVL_CELL_SETTINGS.UNLOAD_MACHINE,
	stMachineStatus := MACHINE_1_FAULT.MachineStatus,
	stRobotStatus := MACHINE_1_FAULT.RobotStatus,
	eRobotTargetPoint := GVL_ROBOT.Diag.eActivePoint,
	xRobotMotionBusy := xMotionBusy,
	Command => GVL_MACHINE.Command[1],
	Status => GVL_MACHINE.Status[1],
	Diag => GVL_MACHINE.Diag[1],
	Error => GVL_MACHINE.Error[1]
);

MACHINE_2.stPoints.eAbove := E_POINT_NAME.MACHINE_2_ABOVE;
MACHINE_2.stPoints.eChuck := E_POINT_NAME.MACHINE_2_CHUCK_POSITION;
MACHINE_2.stPoints.eChuckApproach := E_POINT_NAME.MACHINE_2_CHUCK_APROACH;
MACHINE_2.stPoints.eInside := E_POINT_NAME.MACHINE_2_INSIDE;
MACHINE_2.stPoints.eNone := E_POINT_NAME.NONE;

MACHINE_2(
	RobotResetRecovery := ROBOT.ResetRecovery,
	xResetCancel := GVL_CELL_CONTROL.xStop OR GVL_CELL_CONTROL.xDisable OR GVL_HMI.xRobotStop,
	xTestInitialize := xTestInitializePulse OR xTestAbortActive,
	uiTestInitialState := GVL_HMI.stTestScenario.auiMachineState[2],
	uiTestProductType := GVL_HMI.stTestScenario.auiMachineType[2],
	xExecute := GVL_CELL_MANAGER.Command.axMachineExecute[2],
	xReset := GVL_HMI.axMachineReset[2],
	xResetGlobal := GVL_CELL_CONTROL.xReset,
	xGlobalError := GVL_CELL_CONTROL.xGlobalError,
	xManualMode := GVL_CELL_CONTROL.xManual,
	xIoManual := xIoManualActive,
	xAutomaticUseEnabled := GVL_HMI.axMachineUsed[2],
	xPointsConfigured := axMachinePointsReady[2],
	xSafetyDoorControlEnabled := GVL_CELL_SETTINGS.eTestEnvironment <> E_CELL_TEST_ENVIRONMENT.NORMAL,
	xHmiOpenSafetyDoor := GVL_HMI.axMachineManualSafetyDoorOpen[2],
	xHmiCloseSafetyDoor := GVL_HMI.axMachineManualSafetyDoorClose[2],
	xHmiOpenHatch := GVL_HMI.axMachineManualHatchOpen[2],
	xHmiCloseHatch := GVL_HMI.axMachineManualHatchClose[2],
	xHmiUnlockHatch := GVL_HMI.axMachineManualHatchUnlock[2],
	xHmiLockHatch := GVL_HMI.axMachineManualHatchLock[2],
	xHmiOpenChuck := GVL_HMI.axMachineManualChuckOpen[2],
	xHmiCloseChuck := GVL_HMI.axMachineManualChuckClose[2],
	xHmiEnable := GVL_HMI.axMachineEnable[2],
	xHmiDisable := GVL_HMI.axMachineDisable[2],
	xHmiSetBlank := GVL_HMI.axMachineSetBlank[2],
	xHmiSetDetail := GVL_HMI.axMachineSetDetail[2],
	xHmiAcceptDoor := GVL_HMI.axMachineAcceptDoor[2],
	xHmiRejectDoor := GVL_HMI.axMachineRejectDoor[2],
	xHmiAcceptRunCNC := GVL_HMI.axMachineAcceptRun[2],
	xHmiRejectRunCNC := GVL_HMI.axMachineRejectRun[2],
	xUseHmiCycleTime := GVL_HMI.xUseHmiCycleTime[2],
	tHmiCycleTime := GVL_HMI.tMachineCycleTime[2],
	stTimeouts := MACHINE_2_FAULT.Timeouts,
	stChangeRecipe := GVL_CELL_SETTINGS.CHANGE_MACHINE,
	stLoadRecipe := GVL_CELL_SETTINGS.LOAD_MACHINE,
	stUnloadRecipe := GVL_CELL_SETTINGS.UNLOAD_MACHINE,
	stMachineStatus := MACHINE_2_FAULT.MachineStatus,
	stRobotStatus := MACHINE_2_FAULT.RobotStatus,
	eRobotTargetPoint := GVL_ROBOT.Diag.eActivePoint,
	xRobotMotionBusy := xMotionBusy,
	Command => GVL_MACHINE.Command[2],
	Status => GVL_MACHINE.Status[2],
	Diag => GVL_MACHINE.Diag[2],
	Error => GVL_MACHINE.Error[2]
);

MACHINE_3.stPoints.eAbove := E_POINT_NAME.MACHINE_3_ABOVE;
MACHINE_3.stPoints.eChuck := E_POINT_NAME.MACHINE_3_CHUCK_POSITION;
MACHINE_3.stPoints.eChuckApproach := E_POINT_NAME.MACHINE_3_CHUCK_APROACH;
MACHINE_3.stPoints.eInside := E_POINT_NAME.MACHINE_3_INSIDE;
MACHINE_3.stPoints.eNone := E_POINT_NAME.NONE;

MACHINE_3(
	RobotResetRecovery := ROBOT.ResetRecovery,
	xResetCancel := GVL_CELL_CONTROL.xStop OR GVL_CELL_CONTROL.xDisable OR GVL_HMI.xRobotStop,
	xTestInitialize := xTestInitializePulse OR xTestAbortActive,
	uiTestInitialState := GVL_HMI.stTestScenario.auiMachineState[3],
	uiTestProductType := GVL_HMI.stTestScenario.auiMachineType[3],
	xExecute := GVL_CELL_MANAGER.Command.axMachineExecute[3],
	xReset := GVL_HMI.axMachineReset[3],
	xResetGlobal := GVL_CELL_CONTROL.xReset,
	xGlobalError := GVL_CELL_CONTROL.xGlobalError,
	xManualMode := GVL_CELL_CONTROL.xManual,
	xIoManual := xIoManualActive,
	xAutomaticUseEnabled := GVL_HMI.axMachineUsed[3],
	xPointsConfigured := axMachinePointsReady[3],
	xSafetyDoorControlEnabled := GVL_CELL_SETTINGS.eTestEnvironment <> E_CELL_TEST_ENVIRONMENT.NORMAL,
	xHmiOpenSafetyDoor := GVL_HMI.axMachineManualSafetyDoorOpen[3],
	xHmiCloseSafetyDoor := GVL_HMI.axMachineManualSafetyDoorClose[3],
	xHmiOpenHatch := GVL_HMI.axMachineManualHatchOpen[3],
	xHmiCloseHatch := GVL_HMI.axMachineManualHatchClose[3],
	xHmiUnlockHatch := GVL_HMI.axMachineManualHatchUnlock[3],
	xHmiLockHatch := GVL_HMI.axMachineManualHatchLock[3],
	xHmiOpenChuck := GVL_HMI.axMachineManualChuckOpen[3],
	xHmiCloseChuck := GVL_HMI.axMachineManualChuckClose[3],
	xHmiEnable := GVL_HMI.axMachineEnable[3],
	xHmiDisable := GVL_HMI.axMachineDisable[3],
	xHmiSetBlank := GVL_HMI.axMachineSetBlank[3],
	xHmiSetDetail := GVL_HMI.axMachineSetDetail[3],
	xHmiAcceptDoor := GVL_HMI.axMachineAcceptDoor[3],
	xHmiRejectDoor := GVL_HMI.axMachineRejectDoor[3],
	xHmiAcceptRunCNC := GVL_HMI.axMachineAcceptRun[3],
	xHmiRejectRunCNC := GVL_HMI.axMachineRejectRun[3],
	xUseHmiCycleTime := GVL_HMI.xUseHmiCycleTime[3],
	tHmiCycleTime := GVL_HMI.tMachineCycleTime[3],
	stTimeouts := MACHINE_3_FAULT.Timeouts,
	stChangeRecipe := GVL_CELL_SETTINGS.CHANGE_MACHINE,
	stLoadRecipe := GVL_CELL_SETTINGS.LOAD_MACHINE,
	stUnloadRecipe := GVL_CELL_SETTINGS.UNLOAD_MACHINE,
	stMachineStatus := MACHINE_3_FAULT.MachineStatus,
	stRobotStatus := MACHINE_3_FAULT.RobotStatus,
	eRobotTargetPoint := GVL_ROBOT.Diag.eActivePoint,
	xRobotMotionBusy := xMotionBusy,
	Command => GVL_MACHINE.Command[3],
	Status => GVL_MACHINE.Status[3],
	Diag => GVL_MACHINE.Diag[3],
	Error => GVL_MACHINE.Error[3]
);

// Публичный IO-снимок совпадает с обратной связью, которую анализирует FB_MACHINE.
GVL_MACHINE.Status[1].stIo := MACHINE_1_FAULT.MachineStatus;
GVL_MACHINE.Status[2].stIo := MACHINE_2_FAULT.MachineStatus;
GVL_MACHINE.Status[3].stIo := MACHINE_3_FAULT.MachineStatus;

(* ---- PLC_PRG.RunMagazine.st ---- *)
METHOD PRIVATE RunMagazine

// --- BEGIN IMPLEMENTATION ---

auiMagazineEditSlot[1] := GVL_HMI.astMagazineCommand[1].uiEditSlot;
IF auiMagazineEditSlot[1] = UINT#0 THEN
	auiMagazineEditSlot[1] := GVL_HMI.uiMagazineEditSlot;
END_IF;
auiMagazineEditSlot[2] := GVL_HMI.astMagazineCommand[2].uiEditSlot;

fbMagazine1(
	RobotResetRecovery := ROBOT.ResetRecovery,
	xResetCancel := GVL_CELL_CONTROL.xStop OR GVL_CELL_CONTROL.xDisable OR GVL_HMI.xRobotStop,
	uiMagazineId := UINT#1,
	xInventoryChanged := axMagazineInventoryChanged[1],
	xPointsConfigured := axMagazinePointsReady[1],
	xMechanismReady := (GVL_TWO_PALLET.uiMode = 0) OR GVL_TWO_PALLET.astStatus[1].xReady,
	xTestInitialize := xTestInitializePulse OR xTestAbortActive,
	xTestEnabled := GVL_HMI.stTestScenario.axMagazineEnabled[1],
	stRobotStatus := GVL_ROBOT.Status,
	astMachineStatus := GVL_MACHINE.Status,
	auiMachineType := GVL_MULTI_TYPE.Config.auiMachineType,
	stMagazineCommand := GVL_MAGAZINE.astAutoCommand[1],
	stHmiCommand := GVL_HMI.stRobotCommand,
	xManual := GVL_CELL_CONTROL.xManual AND NOT GVL_CELL_MANAGER.Status.xRunning,
	xIoManual := xIoManualActive,
	xReset := GVL_CELL_CONTROL.xReset OR GVL_HMI.astMagazineCommand[1].xReset OR ((GVL_TWO_PALLET.uiMode = 1) AND (GVL_TWO_PALLET.auiCommand[1] = 16) AND GVL_TWO_PALLET.astStatus[1].xCommandAccepted),
	xGlobalError := GVL_CELL_CONTROL.xGlobalError,
	xHmiEnable := ((GVL_TWO_PALLET.uiMode = 0) AND (GVL_HMI.astMagazineCommand[1].xEnable OR GVL_HMI.xMagazineEnable))
		OR ((GVL_TWO_PALLET.uiMode = 1) AND GVL_TWO_PALLET.astStatus[1].xReady
			AND NOT axTwinMagazineExchangeInProgress[1]
			AND NOT fbMagazine1.Status.xEnabled AND NOT fbMagazine1.Status.xFinished),
	xHmiDisable := GVL_HMI.astMagazineCommand[1].xDisable OR GVL_HMI.xMagazineDisable OR ((GVL_TWO_PALLET.uiMode = 1) AND (NOT GVL_TWO_PALLET.astStatus[1].xEnabled OR GVL_TWO_PALLET.astStatus[1].xBusy OR axTwinMagazineExchangeInProgress[1])),
	xHmiFillBlanks := (GVL_TWO_PALLET.uiMode = 0) AND (GVL_HMI.astMagazineCommand[1].xFill OR GVL_HMI.xMagazineFillBlanks),
	xHmiClear := (GVL_TWO_PALLET.uiMode = 0) AND (GVL_HMI.astMagazineCommand[1].xClear OR GVL_HMI.xMagazineClear),
	xHmiCycleSlot := (GVL_TWO_PALLET.uiMode = 0) AND (GVL_HMI.astMagazineCommand[1].xCycleSlot OR GVL_HMI.xMagazineCycleSlot),
	xHmiApplySlot := (GVL_TWO_PALLET.uiMode = 0) AND (GVL_HMI.astMagazineCommand[1].xApplySlot),
	xHmiApplyPitchX := GVL_HMI.astMagazineCommand[1].xApplyPitchX,
	xHmiApplyPitchY := GVL_HMI.astMagazineCommand[1].xApplyPitchY,
	uiHmiEditSlot := auiMagazineEditSlot[1],
	uiHmiEditDetailType := GVL_HMI.astMagazineCommand[1].uiEditDetailType,
	uiHmiEditProductType := GVL_HMI.astMagazineCommand[1].uiEditProductType,
	lrHmiEditPitchX := GVL_HMI.astMagazineCommand[1].lrEditPitchX,
	lrHmiEditPitchY := GVL_HMI.astMagazineCommand[1].lrEditPitchY,
	xRobotOwnsMagazine := (GVL_CELL_MANAGER.Status.uiActiveMagazine = UINT#1)
		AND (GVL_CELL_MANAGER.Status.xRunning OR GVL_ROBOT.Status.xBusy),
	xRobotCanWorkWithMagazine := xRobotInterfaceReady
		AND axMagazinePointsReady[1]
		AND NOT axTwinMagazineExchangeInProgress[1]
		AND NOT GVL_ROBOT.Status.xError,
	xSharedGeometryEditAllowed := NOT GVL_MAGAZINE.astStatus[1].xEnabled
		AND NOT GVL_MAGAZINE.astStatus[2].xEnabled
		AND NOT GVL_HMI.xMagazineEnable
		AND NOT GVL_HMI.astMagazineCommand[1].xEnable
		AND NOT GVL_HMI.astMagazineCommand[2].xEnable,
	uiRows := GVL_CELL_SETTINGS.MagazineRows,
	uiColumns := GVL_CELL_SETTINGS.MagazineColumns,
	uiTypeCount := GVL_MULTI_TYPE.Config.uiTypeCount,
	auiSlotType := GVL_MULTI_TYPE.Config.auiSlotType,
	FaultRequest := astMagazineFaultRequest[1],
	stInventory := GVL_DETAIL.astMagazine[1],
	lrPitchX := GVL_HMI.MagazinePitchX,
	lrPitchY := GVL_HMI.MagazinePitchY,
	Command => GVL_MAGAZINE.astCommand[1],
	Status => GVL_MAGAZINE.astPartStatus[1],
	Diag => GVL_MAGAZINE.astDiag[1],
	Error => GVL_MAGAZINE.astError[1]
);

fbMagazine2(
	RobotResetRecovery := ROBOT.ResetRecovery,
	xResetCancel := GVL_CELL_CONTROL.xStop OR GVL_CELL_CONTROL.xDisable OR GVL_HMI.xRobotStop,
	uiMagazineId := UINT#2,
	xInventoryChanged := axMagazineInventoryChanged[2],
	xPointsConfigured := axMagazinePointsReady[2],
	xMechanismReady := (GVL_TWO_PALLET.uiMode = 0) OR GVL_TWO_PALLET.astStatus[2].xReady,
	xTestInitialize := xTestInitializePulse OR xTestAbortActive,
	xTestEnabled := GVL_HMI.stTestScenario.axMagazineEnabled[2],
	stRobotStatus := GVL_ROBOT.Status,
	astMachineStatus := GVL_MACHINE.Status,
	auiMachineType := GVL_MULTI_TYPE.Config.auiMachineType,
	stMagazineCommand := GVL_MAGAZINE.astAutoCommand[2],
	stHmiCommand := GVL_HMI.stRobotCommand,
	xManual := GVL_CELL_CONTROL.xManual AND NOT GVL_CELL_MANAGER.Status.xRunning,
	xIoManual := xIoManualActive,
	xReset := GVL_CELL_CONTROL.xReset OR GVL_HMI.astMagazineCommand[2].xReset OR ((GVL_TWO_PALLET.uiMode = 1) AND (GVL_TWO_PALLET.auiCommand[2] = 16) AND GVL_TWO_PALLET.astStatus[2].xCommandAccepted),
	xGlobalError := GVL_CELL_CONTROL.xGlobalError,
	xHmiEnable := ((GVL_TWO_PALLET.uiMode = 0) AND (GVL_HMI.astMagazineCommand[2].xEnable))
		OR ((GVL_TWO_PALLET.uiMode = 1) AND GVL_TWO_PALLET.astStatus[2].xReady
			AND NOT axTwinMagazineExchangeInProgress[2]
			AND NOT fbMagazine2.Status.xEnabled AND NOT fbMagazine2.Status.xFinished),
	xHmiDisable := GVL_HMI.astMagazineCommand[2].xDisable OR ((GVL_TWO_PALLET.uiMode = 1) AND (NOT GVL_TWO_PALLET.astStatus[2].xEnabled OR GVL_TWO_PALLET.astStatus[2].xBusy OR axTwinMagazineExchangeInProgress[2])),
	xHmiFillBlanks := (GVL_TWO_PALLET.uiMode = 0) AND (GVL_HMI.astMagazineCommand[2].xFill),
	xHmiClear := (GVL_TWO_PALLET.uiMode = 0) AND (GVL_HMI.astMagazineCommand[2].xClear),
	xHmiCycleSlot := (GVL_TWO_PALLET.uiMode = 0) AND (GVL_HMI.astMagazineCommand[2].xCycleSlot),
	xHmiApplySlot := (GVL_TWO_PALLET.uiMode = 0) AND (GVL_HMI.astMagazineCommand[2].xApplySlot),
	xHmiApplyPitchX := GVL_HMI.astMagazineCommand[2].xApplyPitchX,
	xHmiApplyPitchY := GVL_HMI.astMagazineCommand[2].xApplyPitchY,
	uiHmiEditSlot := auiMagazineEditSlot[2],
	uiHmiEditDetailType := GVL_HMI.astMagazineCommand[2].uiEditDetailType,
	uiHmiEditProductType := GVL_HMI.astMagazineCommand[2].uiEditProductType,
	lrHmiEditPitchX := GVL_HMI.astMagazineCommand[2].lrEditPitchX,
	lrHmiEditPitchY := GVL_HMI.astMagazineCommand[2].lrEditPitchY,
	xRobotOwnsMagazine := (GVL_CELL_MANAGER.Status.uiActiveMagazine = UINT#2)
		AND (GVL_CELL_MANAGER.Status.xRunning OR GVL_ROBOT.Status.xBusy),
	xRobotCanWorkWithMagazine := xRobotInterfaceReady
		AND axMagazinePointsReady[2]
		AND NOT axTwinMagazineExchangeInProgress[2]
		AND NOT GVL_ROBOT.Status.xError,
	xSharedGeometryEditAllowed := NOT GVL_MAGAZINE.astStatus[1].xEnabled
		AND NOT GVL_MAGAZINE.astStatus[2].xEnabled
		AND NOT GVL_HMI.xMagazineEnable
		AND NOT GVL_HMI.astMagazineCommand[1].xEnable
		AND NOT GVL_HMI.astMagazineCommand[2].xEnable,
	uiRows := GVL_CELL_SETTINGS.MagazineRows,
	uiColumns := GVL_CELL_SETTINGS.MagazineColumns,
	uiTypeCount := GVL_MULTI_TYPE.Config.uiTypeCount,
	auiSlotType := GVL_MULTI_TYPE.Config.auiSlotType,
	FaultRequest := astMagazineFaultRequest[2],
	stInventory := GVL_DETAIL.astMagazine[2],
	lrPitchX := GVL_HMI.MagazinePitchX,
	lrPitchY := GVL_HMI.MagazinePitchY,
	Command => GVL_MAGAZINE.astCommand[2],
	Status => GVL_MAGAZINE.astPartStatus[2],
	Diag => GVL_MAGAZINE.astDiag[2],
	Error => GVL_MAGAZINE.astError[2]
);

// Сохранить физический инвентарь текущей палеты после подтверждённых действий робота.
FOR uiTwin := 1 TO 2 DO
	GVL_MAGAZINE.astStatus[uiTwin] := GVL_MAGAZINE.astPartStatus[uiTwin];
	IF NOT GVL_TWO_PALLET.astStatus[uiTwin].xError THEN axTwinRobotStopLatched[uiTwin] := FALSE;
	ELSIF GVL_ROBOT.Status.uiMagazineContext = uiTwin THEN axTwinRobotStopLatched[uiTwin] := TRUE; END_IF;
	IF GVL_TWO_PALLET.uiMode = 1 THEN
		uiTwinPallet := GVL_TWO_PALLET.astStatus[uiTwin].uiRobotPallet;
		IF (uiTwinPallet >= UINT#1) AND (uiTwinPallet <= UINT#2) THEN
            IF ((uiTwin = UINT#1) AND fbMagazine1.xInventoryUpdated)
            OR ((uiTwin = UINT#2) AND fbMagazine2.xInventoryUpdated) THEN
                GVL_TWO_PALLET.astStore[uiTwin].astPallet[uiTwinPallet] := GVL_DETAIL.astMagazine[uiTwin];
                axTwinStoreChanged[uiTwin] := TRUE;
            END_IF;
		END_IF;
		GVL_MAGAZINE.astStatus[uiTwin].xReady := GVL_MAGAZINE.astStatus[uiTwin].xReady AND GVL_TWO_PALLET.astStatus[uiTwin].xReady;
		GVL_MAGAZINE.astStatus[uiTwin].xEnableSequenceAllowed := GVL_TWO_PALLET.astStatus[uiTwin].xEnableAllowed;
		GVL_MAGAZINE.astStatus[uiTwin].xEnabled := GVL_TWO_PALLET.astStatus[uiTwin].xEnabled;
		GVL_MAGAZINE.astStatus[uiTwin].xBusy := GVL_MAGAZINE.astPartStatus[uiTwin].xBusy OR GVL_TWO_PALLET.astStatus[uiTwin].xBusy;
		GVL_MAGAZINE.astStatus[uiTwin].xFillAllowed := FALSE;
		GVL_MAGAZINE.astStatus[uiTwin].xClearAllowed := FALSE;
		GVL_MAGAZINE.astStatus[uiTwin].xEditAllowed := FALSE;
		GVL_MAGAZINE.astStatus[uiTwin].xError := GVL_MAGAZINE.astStatus[uiTwin].xError OR GVL_TWO_PALLET.astStatus[uiTwin].xError;
		GVL_MAGAZINE.astError[uiTwin].dwErrorActive := GVL_MAGAZINE.astError[uiTwin].dwErrorActive
			OR GVL_TWO_PALLET.astError[uiTwin].dwErrorActive;
		GVL_MAGAZINE.astError[uiTwin].dwAlarmActive := GVL_MAGAZINE.astError[uiTwin].dwAlarmActive
			OR GVL_TWO_PALLET.astError[uiTwin].dwAlarmActive;
		GVL_MAGAZINE.astStatus[uiTwin].xRobotStopRequired := GVL_MAGAZINE.astStatus[uiTwin].xRobotStopRequired
			OR axTwinRobotStopLatched[uiTwin];
		IF axTwinRobotStopLatched[uiTwin] THEN
			GVL_MAGAZINE.astCommand[uiTwin].xStop := TRUE;
			GVL_MAGAZINE.astCommand[uiTwin].xExecute := FALSE;
		END_IF;
	ELSE
        IF ((uiTwin = UINT#1) AND fbMagazine1.xInventoryUpdated)
        OR ((uiTwin = UINT#2) AND fbMagazine2.xInventoryUpdated) THEN
            GVL_TWO_PALLET.astStatic[uiTwin] := GVL_DETAIL.astMagazine[uiTwin];
        END_IF;
	END_IF;
END_FOR;

IF GVL_TWO_PALLET.uiMode = 0 THEN
	Persistent_Value.lrStaticPitchX := GVL_HMI.MagazinePitchX;
	Persistent_Value.lrStaticPitchY := GVL_HMI.MagazinePitchY;
ELSE
	Persistent_Value.lrTwinPitchX := GVL_HMI.MagazinePitchX;
	Persistent_Value.lrTwinPitchY := GVL_HMI.MagazinePitchY;
END_IF;
